	wEncoderID					:WORD := 0; 				(* Encoder ID number *)
	lrTaskCycle					:LREAL := 0.002; 			(* Cycle time of the task which is defined for NC [sec] *)
	bCountDirInv					:BOOL := FALSE;			(* Counting direction inverted if TRUE *)
	udnScalingDenom				:UDINT := 1;	  			(* Denominator for the conversion factor at the conversion of bus data to technical units [INC] *)
	lrScalingNum					:LREAL := 1.0;  			(* Numerator for the conversion factor at the conversion of bus data to technical units [technical units] *)
														(* The technical units dependent on denominator and numerator.*)
	lrModuloFactor 				:LREAL := 360.0; 			(* The "distance" represented by one rotation [technical units] *) 
	dwModuloValue				:DWORD := 0; 			(* Maximum encoder modulo value e.g 1048576 [inc] *)
	etScalingMethod				:ET_ScalingMethod := ET_ScalingMethod_eSMLinear; (* Scaling method: linear or rotary *)
	bSWLimitMaxEn				:BOOL := FALSE;			(* Activation and deactivation of the monitoring of the maximum end position. *)
	lrSWPosLimitMax				:LREAL := 0.0;				(* Location of the maximum end position [technical units] *)
	bSWLimitMinEn 				:BOOL := FALSE;			(* Activation and deactivation of the monitoring of the minimum end position. *)
	lrSWPosLimitMin				:LREAL := 0.0;				(* Location of the minimum end position [technical units] *)

END_STRUCT
END_TYPE

// ---- Data types/Objects/Axis/InternalMC/ST_AXIS_REF_V2.TcDUT
TYPE ST_AXIS_REF_V2 : FB_AXIS_REF_V2;
END_TYPE

// ---- Data types/Objects/EtherCAT Diag/ET_EtherCATDiag.TcDUT
TYPE ET_EtherCATDiag :
(
	ET_EtherCATDiag_eIdle := 0,
	ET_EtherCATDiag_eGetSlaveAdresses,
	ET_EtherCATDiag_eGetSlaveStates,
	ET_EtherCATDiag_eGetTopologyDataLen,
	ET_EtherCATDiag_eGetTopologyData,
	ET_EtherCATDiag_eScanSlaves,
	ET_EtherCATDiag_eGetSlaveIdentity,
	ET_EtherCATDiag_eGetSlaveName,
	ET_EtherCATDiag_eGetScannedSlaveName,
	ET_EtherCATDiag_eDone := 197
);
END_TYPE

// ---- Data types/Objects/EtherCAT Diag/E_EcCommState.TcDUT
TYPE E_EcCommState : (
	eEcState_UNDEFINED 	:= 0,
	eEcState_INIT 		:= 1,
	eEcState_PREOP 		:= 2,
	eEcState_BOOT 		:= 3,
	eEcState_SAFEOP 	:= 4,
	eEcState_OP 		:= 8
);
END_TYPE

// ---- Data types/Objects/EtherCAT Diag/ST_EcMasterDevState.TcDUT
TYPE ST_EcMasterDevState :
STRUCT
	eEcState	 		: E_EcCommState;
	nReserved			: ARRAY [0..2] OF UINT;

	bLinkError			: BOOL;
	bResetRequired		: BOOL;
	bMissFrmRedMode		: BOOL;
	bWatchdogTriggerd	: BOOL;
	bDriverNotFound		: BOOL;
	bResetActive		: BOOL;
	bAtLeastOneNotInOp	: BOOL;
	bDcNotInSync		: BOOL;
END_STRUCT
END_TYPE

// ---- Data types/Objects/EtherCAT Diag/ST_SlaveState.TcDUT
TYPE ST_SlaveState :
STRUCT
	(* slave state *)
	eEcState 		: E_EcCommState;
	nReserved		: UINT;
	bError			: BOOL;
	bInvalidVPRS	: BOOL;
	nReserved2		: UINT;

	(* link state *)
	bNoCommToSlave	: BOOL;
	bLinkError		: BOOL;
	bMissingLink	: BOOL;
	bUnexpectedLink	: BOOL;
	bPortA			: BOOL;
	bPortB			: BOOL;
	bPortC			: BOOL;
	bPortD			: BOOL;
END_STRUCT
END_TYPE

// ---- Data types/Objects/EtherCAT Diag/ST_SlaveStateInfo.TcDUT
TYPE ST_SlaveStateInfo :
STRUCT
	nIndex 			: DINT;
	sName 			: STRING; 		(* name of slave given in System Manager *)
	sType 			: STRING;		(* type of slave, e.g. EK1100*)
	nECAddr 		: UINT;			(* EtherCAT Slave Addr *)
	bDiagData		: BOOL;			(* DiagData in Slave State *)
	stPortCRCErrors	: ST_EcCrcErrorEx;(* Slave CRC-Errors, separate for each Port *)
	nSumCRCErrors	: UDINT;		(* Slave CRC-Errors, sum of all Ports *)
	stState 		: ST_SlaveState;(* EtherCAT State and Link state*)
END_STRUCT
END_TYPE

// ---- Data types/Objects/EtherCAT Diag/ST_SlaveStateInfoScanned.TcDUT
TYPE ST_SlaveStateInfoScanned :
STRUCT
	nIndex 			: DINT;
	sName 			: STRING; 		(* name of slave given in System Manager *)
	sType 			: STRING;		(* type of slave, e.g. EK1100*)
	nECAddr 		: UINT;			(* EtherCAT Slave Addr *)
	bDifferentName	: BOOL;			(* Name of Scanned configuration differs from Configured configuration *)
	bDifferentType	: BOOL;			(* Type Of Scanned configuration differs from Configured configuration *)
	bDifferentAddr	: BOOL;			(* EcAddress of Scanned configuration differs from Configured configuration *)
END_STRUCT
END_TYPE

// ---- Data types/Objects/EtherCAT Diag/ST_TopologyData.TcDUT
TYPE ST_TopologyData :
STRUCT
	iOwnPhysicalAddr 	: UINT;
	iOwnAutoIncAddr		: UINT;
	stPhysicalAddr		: ST_PortAddr;
	stAutoIncAddr		: ST_PortAddr;
	iPortDelay			: ARRAY [0..2] OF UDINT; (* EC_AD, EC_DB, EC_BC *)
	iReserved			: ARRAY [0..7] OF UDINT;
END_STRUCT
END_TYPE

// ---- Data types/Objects/ET_SpindleCtrl/ET_SpindleCtrl.TcDUT
TYPE ET_SpindleCtrl :
(
	ET_SpindleCtrl_eWaitExecute := 0,
	ET_SpindleCtrl_eCtrlEnable := 5,
	ET_SpindleCtrl_eWfCtrlEnabled := 10,
	ET_SpindleCtrl_eSpindleStop := 15,
	ET_SpindleCtrl_eWfSpindleStopped := 20,
	ET_SpindleCtrl_eSpindleRun := 25,
	ET_SpindleCtrl_eWfSpindleRunning := 30,
	ET_SpindleCtrl_eDone := 197,
	ET_SpindleCtrl_eError := 198,
	ET_SpindleCtrl_eNoExecute := 199
);
END_TYPE

// ---- Data types/Objects/FB_Alarm/ET_AlarmType.TcDUT
TYPE ET_AlarmType :
(
	ET_AlarmType_eIdle := 0,
	ET_AlarmType_eFatalError := 1,
	ET_AlarmType_eError := 2,
	ET_AlarmType_eWarning := 3,
	ET_AlarmType_eMessage := 4,
	ET_AlarmType_eHint := 5
);
END_TYPE

// ---- Data types/Objects/FB_Alarm/ST_Alarm.TcDUT
TYPE ST_Alarm :
STRUCT
	bFatalError			:BOOL;				(* Fatal error in group / Fataler Fehler in der Gruppe *)
	bError				:BOOL;				(* Error in group / Fehler in der Gruppe *)
	bWarning			:BOOL;				(* Warning in group / Warnung  in der Gruppe *)
	bMessage			:BOOL;				(* Message in group / Meldung in der Gruppe *)
	bHint				:BOOL;				(* Hint in group / Hint in der Gruppe *)
END_STRUCT
END_TYPE

// ---- Data types/Objects/FB_Alarm/ST_AlarmIn.TcDUT
TYPE ST_AlarmIn :
STRUCT
	arbFatalError			:ARRAY[0..nALARM_MAX_NO] OF ST_AlarmProperties;
	arbError				:ARRAY[0..nALARM_MAX_NO] OF ST_AlarmProperties;
	arbWarning			:ARRAY[0..nALARM_MAX_NO] OF ST_AlarmProperties;
	arbMessage			:ARRAY[0..nALARM_MAX_NO] OF ST_AlarmProperties;
	arbHint				:ARRAY[0..nALARM_MAX_NO] OF ST_AlarmProperties;
END_STRUCT
END_TYPE

// ---- Data types/Objects/FB_Alarm/ST_AlarmOut.TcDUT
TYPE ST_AlarmOut :
STRUCT
	arbFatalError			:ARRAY[0..nALARM_MAX_NO] OF ST_AlarmProperties;
	arbError				:ARRAY[0..nALARM_MAX_NO] OF ST_AlarmProperties;
	arbWarning			:ARRAY[0..nALARM_MAX_NO] OF ST_AlarmProperties;
	arbMessage			:ARRAY[0..nALARM_MAX_NO] OF ST_AlarmProperties;
	arbHint				:ARRAY[0..nALARM_MAX_NO] OF ST_AlarmProperties;
	bFatalError			:BOOL;				(* Fatal error in group / Fataler Fehler in der Gruppe *)
	bError				:BOOL;				(* Error in group / Fehler in der Gruppe *)
	bWarning			:BOOL;				(* Warning in group / Warnung  in der Gruppe *)
	bMessage			:BOOL;				(* Message in group / Meldung in der Gruppe *)
	bHint				:BOOL;				(* Hint in group / Hint in der Gruppe *)
END_STRUCT
END_TYPE

// ---- Data types/Objects/FB_Alarm/ST_AlarmProperties.TcDUT
TYPE ST_AlarmProperties :
STRUCT
	bActive				:BOOL;				(* Alarm on *)
	dtDateTime			:DATE_AND_TIME ;	(* Alarm time stamp *)
	enType				:ET_AlarmType;		(* Alarm type *)
	dnCode				:DINT;				(* Alarm code *)
END_STRUCT
END_TYPE

// ---- Data types/Objects/FB_Alarm/ST_AlarmRef.TcDUT
TYPE ST_AlarmRef :
STRUCT
	stControl					:ST_AlarmOut;
	stManual					:ST_AlarmOut;
	stMaintenance			:ST_AlarmOut;
	stHome					:ST_AlarmOut;
	stAuto					:ST_AlarmOut;
END_STRUCT
END_TYPE

// ---- Data types/Objects/FB_AxisController/ET_AxisGetLimits.TcDUT
TYPE ET_AxisGetLimits :
(
	ET_AxisGetLimits_eWaitExecute := 0,
	ET_AxisGetLimits_eReadVeloMax,
	ET_AxisGetLimits_eWfReadVeloMax,
	ET_AxisGetLimits_eReadAccMax,
	ET_AxisGetLimits_eWfReadAccMax,
	ET_AxisGetLimits_eReadDecMax,
	ET_AxisGetLimits_eWfReadDecMax,
	ET_AxisGetLimits_eReadJerkMax,
	ET_AxisGetLimits_eWfReadJerkMax,
	ET_AxisGetLimits_eReadSoftLimitMax,
	ET_AxisGetLimits_eWfReadSoftLimitMax,
	ET_AxisGetLimits_eReadSoftLimitMin,
	ET_AxisGetLimits_eWfReadSoftLimitMin,
	ET_AxisGetLimits_eDone := 197,
	ET_AxisGetLimits_eError := 198,
	ET_AxisGetLimits_eNoExecute := 199
);
END_TYPE

// ---- Data types/Objects/FB_AxisController/ET_AxisSetLimits.TcDUT
TYPE ET_AxisSetLimits :
(
	ET_AxisSetLimits_eWaitExecute := 0,
	ET_AxisSetLimits_eSetReferenceSystem,
	ET_AxisSetLimits_eWfSetReferenceSystem,
	ET_AxisSetLimits_eSetPositionBias,
	ET_AxisSetLimits_eWfSetPositionBias,
	ET_AxisSetLimits_eSetLimitPos,
	ET_AxisSetLimits_eWfSetLimitPos,
	ET_AxisSetLimits_eSetLimitNeg,
	ET_AxisSetLimits_eWfSetLimitNeg,
	ET_AxisSetLimits_eEnableLimitPos,
	ET_AxisSetLimits_eWfEnableLimitPos,
	ET_AxisSetLimits_eEnableLimitNeg,
	ET_AxisSetLimits_eWfEnableLimitNeg,
	ET_AxisSetLimits_eEnablePosLagMonitoring,
	ET_AxisSetLimits_eWfEnablePosLagMonitoring,
	ET_AxisSetLimits_eDone := 197,
	ET_AxisSetLimits_eError := 198,
	ET_AxisSetLimits_eNoExecute := 199
);
END_TYPE

// ---- Data types/Objects/FB_AxisController/ET_STOEBER_AxisGetLimitsTc2.TcDUT
TYPE ET_STOEBER_AxisGetLimitsTc2 :
(
	ET_STOEBER_AxisGetLimits_eWaitExecute := 0,
	ET_STOEBER_AxisGetLimits_eDecimalDigits,
	ET_STOEBER_AxisGetLimits_eScalingDenom,
	ET_STOEBER_AxisGetLimits_eScalingNum,
	ET_STOEBER_AxisGetLimits_eDone := 197,
	ET_STOEBER_AxisGetLimits_eError := 198,
	ET_STOEBER_AxisGetLimits_eNoExecute := 199
);
END_TYPE

// ---- Data types/Objects/FB_AxisController/ET_STOEBER_AxisSetLimitsTc2.TcDUT
TYPE ET_STOEBER_AxisSetLimitsTc2 :
(
	ET_STOEBER_AxisSetLimits_eWaitExecute := 0,
	ET_STOEBER_AxisSetLimits_eSetLimitPos,
	ET_STOEBER_AxisSetLimits_eSetLimitNeg,
	ET_STOEBER_AxisSetLimits_eSetJogVelo,
	ET_STOEBER_AxisSetLimits_eSetJogAcc,
	ET_STOEBER_AxisSetLimits_eSetJogDec,
	ET_STOEBER_AxisSetLimits_eSetJogJerk,
	ET_STOEBER_AxisSetLimits_eDone := 197,
	ET_STOEBER_AxisSetLimits_eError := 198,
	ET_STOEBER_AxisSetLimits_eNoExecute := 199
);
END_TYPE

// ---- Data types/Objects/FB_AxisMoveManual/ET_AxisMoveManualSetLimits.TcDUT
TYPE ET_AxisMoveManualSetLimits :
(
	ET_AxisMoveManualSetLimits_eWaitExecute := 0,
	ET_AxisMoveManualSetLimits_eSetVelo := 5,
	ET_AxisMoveManualSetLimits_eWfSetVelo := 10,
	ET_AxisMoveManualSetLimits_eDone := 197,
	ET_AxisMoveManualSetLimits_eError := 198,
	ET_AxisMoveManualSetLimits_eNoExecute := 199
);
END_TYPE

// ---- Data types/Objects/FB_Blinker/ST_Blinker.TcDUT
TYPE ST_Blinker :
STRUCT	
	Q0					:BOOL; 						(* Divider output / 2 *)
	Q1					:BOOL; 						(* Divider output / 4 *)
	Q2					:BOOL; 						(* Divider output / 8 *)
	Q3					:BOOL; 						(* Divider output / 16 *)
	Q4					:BOOL; 						(* Divider output / 32 *)
	Q5					:BOOL; 						(* Divider output / 64 *)
	Q6					:BOOL; 						(* Divider output / 128 *)
	Q7					:BOOL; 						(* Divider output / 256 *)
END_STRUCT
END_TYPE

// ---- Data types/Objects/FB_CalcContour/ET_ContourType.TcDUT
TYPE ET_ContourType :
(
	ET_ContourType_eNone := 0,
	ET_ContourType_eCircle := 1,
	ET_ContourType_eEllipse := 2,
	ET_ContourType_eSquare := 3
);
END_TYPE

// ---- Data types/Objects/FB_CfgAxisInExt3DGroup/ET_CfgAxisInExt3DGroup.TcDUT
TYPE ET_CfgAxisInExt3DGroup :
(
	ET_CfgAxisInExt3DGrp_eWaitExecute := 0,
	ET_CfgAxisInExt3DGrp_eReadExt3DAxisIds := 5,
	ET_CfgAxisInExt3DGrp_eDone := 197,
	ET_CfgAxisInExt3DGrp_eError := 198,
	ET_CfgAxisInExt3DGrp_eNoExecute := 199
);
END_TYPE

// ---- Data types/Objects/FB_DistanceCounter/ST_DistanceCounter.TcDUT
TYPE ST_DistanceCounter :
STRUCT
	lrAllOverDistance					:LREAL; 							(* All over counter distance *)
	lrAfterResetDistance				:LREAL; 							(* Counter distance since last reset *)
END_STRUCT
END_TYPE

// ---- Data types/Objects/FB_EL3312/ET_EL3312ThermocoupleTyp.TcDUT
TYPE ET_EL3312ThermocoupleTyp :
(
	ET_EL3312ThermocoupleTyp_eK := 0,				(* Typ: K -200°C bis 1370°C *)
	ET_EL3312ThermocoupleTyp_eJ := 1,				(* Typ: J -100°C bis 1200°C *)
	ET_EL3312ThermocoupleTyp_eL := 2,				(* Typ: L 0°C bis 900°C *)
	ET_EL3312ThermocoupleTyp_eE := 3,				(* Typ: E -100°C bis 1000°C *)
	ET_EL3312ThermocoupleTyp_eT := 4,				(* Typ: T -200°C bis 400°C *)
	ET_EL3312ThermocoupleTyp_eN := 5,				(* Typ: N -100°C bis 1300°C *)
	ET_EL3312ThermocoupleTyp_eU := 6,				(* Typ: U 0°C bis 600°C *)
	ET_EL3312ThermocoupleTyp_eB := 7,				(* Typ: B 600°C bis 1800°C *)
	ET_EL3312ThermocoupleTyp_eR := 8,				(* Typ: R 0°C bis 1767°C *)
	ET_EL3312ThermocoupleTyp_eS := 9,				(* Typ: S 0°C bis 1760°C *)
	ET_EL3312ThermocoupleTyp_eC := 10,				(* Typ: C 0°C bis 2320°C *)
	ET_EL3312ThermocoupleTyp_e30mV := 100,			(* +/-30 mV (1uV resolution) *)
	ET_EL3312ThermocoupleTyp_e60mV := 101,			(* +/-60 mV (2uV resolution) *)
	ET_EL3312ThermocoupleTyp_e75mV := 102,			(* +/-75 mV (4uV resolution) *)
	ET_EL3312ThermocoupleTyp_eNoConn := 999		(* No connected *)
);
END_TYPE

// ---- Data types/Objects/FB_EL3312/ST_EL3312ChannelState.TcDUT
TYPE ST_EL3312ChannelState :
STRUCT
	bUnderrange				:BOOL;			(* State underrange *)
	bOverrange				:BOOL;			(* State overrange *)
	byLimit1					:BYTE;			(* State limit 1 *)
	byLimit2 					:BYTE;			(* State limit 2 *)
	bError 					:BOOL;			(* State error *)
	bState 					:BOOL;			(* State *)
	bToggle					:BOOL;			(* TxPDO Toggle *)
END_STRUCT
END_TYPE

// ---- Data types/Objects/FB_EL3312/ST_EL3312CoeInfo.TcDUT
TYPE ST_EL3312CoeInfo :
STRUCT
	bEnableUserScale 			:BOOL := FALSE;
	bEnableFilter 					:BOOL := FALSE;
	bEnableLimit1 				:BOOL := FALSE;
	bEnableLimit2 				:BOOL := FALSE;
	bEnableUserCalibration 		:BOOL := FALSE;
	bEnableVendorCalibration 		:BOOL := TRUE;
	dwColdjunctionCompensation 	:DWORD := 0;
	nUserScaleOffset 				:INT := 0;
	dnUserScaleGain 				:DINT := 65536;
	nLimit1 						:INT := 0;
	nLimit2 						:INT := 0;
	dwFilterSettings 				:DWORD := 0;
	nUserCalibrationOffset 			:INT := 0;
	unUserCalibrationGain 			:UINT := 65535;
	dwTCElement 				:DWORD := 0;
END_STRUCT
END_TYPE

// ---- Data types/Objects/FB_EL3312/ST_EL3312CoeReadData.TcDUT
TYPE ST_EL3312CoeReadData :
STRUCT
	wIdx: WORD;
	bySubIdx: BYTE;
	bReadOK: BOOL;
	dwData: DWORD;
	nSize: UDINT;
END_STRUCT
END_TYPE

// ---- Data types/Objects/FB_EL3312/ST_EL3312CoeWriteData.TcDUT
TYPE ST_EL3312CoeWriteData :
STRUCT
	wIdx: WORD;
	bySubIdx: BYTE;
	bWriteOK: BOOL;
	dwData: DWORD;
	nSize: UDINT;
END_STRUCT
END_TYPE

// ---- Data types/Objects/FB_EL3351/ST_EL3351ChannelState.TcDUT
TYPE ST_EL3351ChannelState :
STRUCT
	bUnderrange				:BOOL;			(* State underrange *)
	bOverrangerange			:BOOL;			(* State overrangerange *)
	bError 					:BOOL;			(* State error *)
	bState 					:BOOL;			(* State *)
	bToggle					:BOOL;			(* TxPDO Toggle *)
END_STRUCT
END_TYPE

// ---- Data types/Objects/FB_EL3351/ST_EL3351CoeInfo.TcDUT
TYPE ST_EL3351CoeInfo :
STRUCT
	bEnableUserScale: BOOL:= 0;
	diUserScaleOffset: DINT:= 0;
	diUserScaleGain: DINT:= 65536;
	dwFilterSettings: DWORD:= 2;

	bEnableUserScaleIndex8010: BOOL:= 0;
	dnUserScaleOffsetIndex8010: DINT:= 0;
	dnUserScaleGainIndex8010: DINT:= 65536;
END_STRUCT
END_TYPE

// ---- Data types/Objects/FB_EL3351/ST_EL3351CoeReadData.TcDUT
TYPE ST_EL3351CoeReadData :
STRUCT
	wIdx: WORD;
	bySubIdx: BYTE;
	bReadOK: BOOL;
	nData: UDINT;
	nSize: UDINT;
END_STRUCT
END_TYPE

// ---- Data types/Objects/FB_EL3351/ST_EL3351CoeWriteData.TcDUT
TYPE ST_EL3351CoeWriteData :
STRUCT
	wIdx: WORD;
	bySubIdx: BYTE;
	bWriteOK: BOOL;
	nData: DWORD;
	nSize: UDINT;
END_STRUCT
END_TYPE

// ---- Data types/Objects/FB_EL3356/ST_EL3356ChannelCtrl.TcDUT
TYPE ST_EL3356ChannelCtrl :
STRUCT
	bStartCalibration			:BOOL;			(* Ctrl start calibration *)
	bDisableCalibration		:BOOL;			(* Ctrl disable calibration *)
	bInputFreeze				:BOOL;			(* Ctrl input freeze *)
	bTare					:BOOL;			(* Ctrl tare *)
END_STRUCT
END_TYPE

// ---- Data types/Objects/FB_EL3356/ST_EL3356ChannelState.TcDUT
TYPE ST_EL3356ChannelState :
STRUCT
	bOverrange				:BOOL;			(* State Overrange *)
	bDataInvalid				:BOOL;			(* State Data invalid *)
	bError 					:BOOL;			(* State error *)
	bCalibrationInProgress 	:BOOL;			(* State calibration in progress *)
	bSteadyState 			:BOOL;			(* Stady state *)
	bSyncError				:BOOL;			(* Sync error *)
	bToggle					:BOOL;			(* TxPDO Toggle *)
END_STRUCT
END_TYPE

// ---- Data types/Objects/FB_EL3356/ST_EL3356CoeInfo.TcDUT
TYPE ST_EL3356CoeInfo :
STRUCT
	bEnableFilter							:BOOL:= TRUE;
	bEnableUserScale					:BOOL:= TRUE;
	dwFilterSettings						:DWORD:= 0;
	rGain								:REAL:= 1.0;
	rTara								:REAL:= 0.0;
	rRatedOutput							:REAL:= 2.0;
	rNominalLoad						:REAL:= 5.0;
	rZeroBalance							:REAL:= 0.0;
	rGravityOfEarth						:REAL:= 9.806650;
	rScaleFactor							:REAL:= 1000.0;
	rReferenceLoad						:REAL:= 5.0;
	bEnableUserScaleIndex8010			:BOOL:= FALSE;
	dnUserScaleOffsetIndex8010			:DINT:= 0;
	dnUserScaleGainIndex8010				:DINT:= 65536;
	dwFilterSettingsIndex8010				:DWORD:= 0;
END_STRUCT
END_TYPE

// ---- Data types/Objects/FB_EL3356/ST_EL3356CoeReadData.TcDUT
TYPE ST_EL3356CoeReadData :
STRUCT
	wIdx: WORD;
	bySubIdx: BYTE;
	bReadOK: BOOL;
	dwData: DWORD;
	nSize: UDINT;
END_STRUCT
END_TYPE

// ---- Data types/Objects/FB_EL3356/ST_EL3356CoeWriteData.TcDUT
TYPE ST_EL3356CoeWriteData :
STRUCT
	wIdx: WORD;
	bySubIdx: BYTE;
	bWriteOK: BOOL;
	dwData: DWORD;
	nSize: UDINT;
END_STRUCT
END_TYPE

// ---- Data types/Objects/FB_ExtSetPoint/ET_MoveExtState.TcDUT
TYPE ET_MoveExtState :
(
	ET_MoveExtState_eWaitExecute := 0,
	ET_MoveExtState_eEnableExtSetPointGenerator := 5,
	ET_MoveExtState_eDisableExtSetPointGenerator := 10,
	ET_MoveExtState_eDone := 197,
	ET_MoveExtState_eError := 198,
	ET_MoveExtState_eNoExecute := 199
);
END_TYPE

// ---- Data types/Objects/FB_ExtTrajPos/ET_CalcExtTrajState.TcDUT
TYPE ET_CalcExtTrajState :
(
	ET_CalcExtTrajState_eWaitExecute := 0,
	ET_CalcExtTrajState_eCalcTrajPos := 5,
	ET_CalcExtTrajState_eDone := 197,
	ET_CalcExtTrajState_eError := 198,
	ET_CalcExtTrajState_eNoExecute := 199
);
END_TYPE

// ---- Data types/Objects/FB_ItpReadRParams/ET_ItpReadRParams.TcDUT
TYPE ET_ItpReadRParams :
(
	ET_ItpReadRParams_eWaitExecute := 0,
	ET_ItpReadRParams_eReadRParams := 5,
	ET_ItpReadRParams_eDone := 197,
	ET_ItpReadRParams_eError := 198,
	ET_ItpReadRParams_eNoExecute := 199
);
END_TYPE

// ---- Data types/Objects/FB_ItpWriteRParams/ET_ItpWriteRParams.TcDUT
TYPE ET_ItpWriteRParams :
(
	ET_ItpWriteRParams_eWaitExecute := 0,
	ET_ItpWriteRParams_eWriteRParams := 5,
	ET_ItpWriteRParams_eDone := 197,
	ET_ItpWriteRParams_eError := 198,
	ET_ItpWriteRParams_eNoExecute := 199
);
END_TYPE

// ---- Data types/Objects/FB_KL600x/ET_KL600xInit.TcDUT
TYPE ET_KL600xInit :
(
	ET_KL600xInit_eInit := 0,
	ET_KL600xInit_eChkSettings,
	ET_KL600xInit_eWriteEnableRTSCTS,
	ET_KL600xInit_eWriteBaudRate,
	ET_KL600xInit_eWriteDataFrame,
	ET_KL600xInit_eDone := 197,
	ET_KL600xInit_eError := 198,
	ET_KL600xInit_eNoExecute := 199
);
END_TYPE

// ---- Data types/Objects/FB_KL600x/ET_KL600xSend.TcDUT
TYPE ET_KL600xSend :
(
	ET_KL600xSend_eInit := 0,
	ET_KL600xSend_eSend,
	ET_KL600xSend_eDone := 197,
	ET_KL600xSend_eError := 198,
	ET_KL600xSend_eNoExecute := 199
);
END_TYPE

// ---- Data types/Objects/FB_KL600x/ST_KL600xData.TcDUT
TYPE ST_KL600xData :
STRUCT
	sDateTime			:STRING;
	sData				:STRING;
END_STRUCT
END_TYPE

// ---- Data types/Objects/FB_LoadFromFile/ET_LoadFromFile.TcDUT

TYPE ET_LoadFromFile :
(
	ET_LoadFromFile_eWaitExecute := 0,
	ET_LoadFromFile_eFileName,
	ET_LoadFromFile_eChkFileExist,
	ET_LoadFromFile_eFileOpen,
	ET_LoadFromFile_eChkFileOpen,
	ET_LoadFromFile_eReadData,
	ET_LoadFromFile_eChkReadData,
	ET_LoadFromFile_eFileClose,
	ET_LoadFromFile_eChkFileClose,
	ET_LoadFromFile_eDone := 197,
	ET_LoadFromFile_eError := 198,
	ET_LoadFromFile_eNoExecute := 199
);
END_TYPE

// ---- Data types/Objects/FB_Logger/ST_Logger.TcDUT
TYPE ST_Logger :
STRUCT
	arstLoggerWaitInterrupt					:ARRAY[1..unLOG_BEFOR_MAX_NO] OF ST_LoggerVar;
	arstLoggerDuringInterrupt				:ARRAY[1..unLOG_DURING_MAX_NO] OF ST_LoggerVar;
	arstLoggerAfterInterrupt					:ARRAY[1..unLOG_AFTER_MAX_NO] OF ST_LoggerVar;
END_STRUCT
END_TYPE

// ---- Data types/Objects/FB_Logger/ST_LoggerVar.TcDUT
TYPE ST_LoggerVar :
STRUCT
	udnCycleNo		:UDINT;
	sTimeStamp		:STRING(15);			(* Alarm time stamp *)
	arsLogVars		:ARRAY[1..unNUM_OF_LOG_VAR] OF STRING(10);
END_STRUCT
END_TYPE

// ---- Data types/Objects/FB_ModeSelector/ET_MachineMode.TcDUT
(* Machine operating mode *)
TYPE ET_MachineMode :
(
	ET_MachineMode_eUndefined := 0,
	ET_MachineMode_eAutomatic := 1,
	ET_MachineMode_eCycle := 2,
	ET_MachineMode_eStepping := 3,
	ET_MachineMode_eHome := 4,
	ET_MachineMode_eManual := 5,
	ET_MachineMode_eMaintenance := 6,
	ET_MachineMode_eDryRun := 7,
	ET_MachineMode_eMDI := 8,
	ET_MachineMode_eIdle := 10
);
END_TYPE

// ---- Data types/Objects/FB_ModeSelector/ET_MachineState.TcDUT
(* Machine state *)
TYPE ET_MachineState :
(
	ET_MachineState_eUndefined := 0,
	ET_MachineState_eAutoExe := 1,
	ET_MachineState_eAutoSteppingExe := 2,
	ET_MachineState_eAutoSteppingNoExe := 3,
	ET_MachineState_eHomeExe := 4,
	ET_MachineState_eHomeRefExe := 5,
	ET_MachineState_eMaintenanceExe := 6,
	ET_MachineState_eIdle := 10
) ;
END_TYPE

// ---- Data types/Objects/FB_RampDirector/ET_RampGenerator.TcDUT
TYPE ET_RampGenerator :
(
	ET_RampGenerator_eWaitExecute := 0,
	ET_RampGenerator_eRunning := 5,
	ET_RampGenerator_eWaiting := 10,
	ET_RampGenerator_eDone := 197,
	ET_RampGenerator_eError := 198,
	ET_RampGenerator_eNotExecute := 199
);
END_TYPE

// ---- Data types/Objects/FB_SpindlePreheat/ET_SpindlePreheat.TcDUT
TYPE ET_SpindlePreheat :
(
	ET_SpindlePreheat_eWaitExecute := 0,
	ET_SpindlePreheat_eStartNewSpindle := 5,
	ET_SpindlePreheat_eStartDailyPreheat := 10,
	ET_SpindlePreheat_eStartSpindle := 15,
	ET_SpindlePreheat_eWfStartSpindle := 20,
	ET_SpindlePreheat_eWfStartSpindleProc := 25,
	ET_SpindlePreheat_eSpindleStop := 30,
	ET_SpindlePreheat_eWfSpindleStopped := 35,
	ET_SpindlePreheat_eDone := 197,
	ET_SpindlePreheat_eError := 198,
	ET_SpindlePreheat_eNoExecute := 199
);
END_TYPE

// ---- Data types/Objects/FB_SpindlePreheat/ST_SpindlePreheat.TcDUT
TYPE ST_SpindlePreheat :
STRUCT
	dwOverride				:DWORD;			(* Override is percent of total speed of spindle. The range of override is from 0%  to 100 %  of rated speed.*)
	tDuration					:TIME;				(* Duration time for current phase *)
	dwSpeedRpm			:DWORD;			(* Current speed RPM - Read Only *)
	otstDuration				:OTSTRUCT;			(* Duration time in OTSTRUCT - Read Only*)
END_STRUCT
END_TYPE

// ---- Data types/Objects/FB_TimeHoursCounter/ST_TimeHoursCounter.TcDUT
TYPE ST_TimeHoursCounter :
STRUCT
	lrAllOverHours					:LREAL; 							(* All over counter hours *)
	lrAfterResetHours					:LREAL; 							(* Counter hours since last reset *)
END_STRUCT
END_TYPE

// ---- Data types/Objects/FB_Timer/ST_DateTime.TcDUT
TYPE ST_DateTime :
STRUCT
	sDate						:STRING;					(* Current data *)
	sTime						:STRING;					(* Current time *)
	sTimeEx						:STRING;					(* Current time extend *)
	sDateTime					:STRING;					(* Current data and time *)
	dtDateTime					:DATE_AND_TIME;				(* Current data and time *)
	sDateTimeEx					:STRING;					(* Current data and time extend *)
	dtDateTimeEx				:DATE_AND_TIME;				(* Current data and time extend *)
END_STRUCT
END_TYPE

// ---- Data types/Objects/FB_Timer/ST_Time.TcDUT
TYPE ST_Time :
STRUCT
	dwSec				:DWORD; 						(* Time in 1 [s] *)
	dwDeciSec			:DWORD; 						(* Time in deci 0.1 [s] *)
	dwCentiSec			:DWORD; 						(* Time in centi 0.01 [s] *)
	dwMiliSec			:DWORD; 						(* Time in mili 0.001 [s] *)
END_STRUCT
END_TYPE

// ---- Data types/Objects/FB_ToolStorage/ET_ToolStatus.TcDUT
TYPE ET_ToolStatus :
(
	ET_ToolStatus_eOk,
	ET_ToolStatus_eNOk,
	ET_ToolStatus_eLifettimeExceeded
);
END_TYPE

// ---- Data types/Objects/FB_ToolStorage/ET_ToolStorage.TcDUT
TYPE ET_ToolStorage :
(
	ET_ToolStorage_eWaitExecute := 0,
	ET_ToolStorage_eGetNewToolNest,
	ET_ToolStorage_eGetOldToolNest,
	ET_ToolStorage_eChkToolPlace,
	ET_ToolStorage_eChkToolPickUp,
	ET_ToolStorage_eDone := 197,
	ET_ToolStorage_eError := 198,
	ET_ToolStorage_eNoExecute := 199
);
END_TYPE

// ---- Data types/Objects/FB_Traceability/ST_Traceability.TcDUT
TYPE ST_Traceability :
STRUCT
	sDateTime				:STRING(15);
	stSettings				:ST_TraceabilitySettings;
	arstData					:ARRAY[1..udnTraceSampleMax,1..udnTraceDataMax] OF ST_TraceabilityData;
END_STRUCT
END_TYPE

// ---- Data types/Objects/FB_Traceability/ST_TraceabilityData.TcDUT
TYPE ST_TraceabilityData :
STRUCT
	sName					:STRING(15);
	sValue					:STRING(15);
	sUnit					:STRING(5);
END_STRUCT
END_TYPE

// ---- Data types/Objects/FB_Traceability/ST_TraceabilitySettings.TcDUT
TYPE ST_TraceabilitySettings :
STRUCT
	sPath								:STRING;						(* Path to file e.g. 'c:\', Hard Disk\ *)
	sFileName							:STRING(20);						(* Name of file *)
	sFileExtension						:STRING(5);						(* File extension  *)
END_STRUCT
END_TYPE

// ---- Data types/Objects/Fieldbus/ST_FieldbusStatus.TcDUT
TYPE ST_FieldbusStatus :
STRUCT
	wFrmXWcState				:WORD; (* link to task related ethercat frame state FrmXWcState *)
	nMasterDeviceId				:UINT;
	nMasterSlaveCount			:UINT;
	nMasterDevState				:UINT;
	arrMasterNetId				:T_AmsNetIdArr;
	nMasterSlaveCountCfg			:UINT;
END_STRUCT
END_TYPE

// ---- Data types/Objects/Gefran/ET_GFX4IR.TcDUT
TYPE ET_GFX4IR :
(
	ET_GFX4IRState_eWaitExecute := 0,
	ET_GFX4IRState_eCtrlOn,
	ET_GFX4IRState_eCtrlOff,
	ET_GFX4IRState_eDone := 197,
	ET_GFX4IRState_eError := 198,
	ET_GFX4IRState_eNoExecute := 199
);
END_TYPE

// ---- Data types/Objects/Gefran/ST_GFX4IRTOPLC.TcDUT
TYPE ST_GFX4IRTOPLC:
STRUCT
	nProcessVariable			:INT;
	wControllerStatus			:WORD;
	nOutputPower				:INT;
	wAmmeterInputOn			:WORD;
END_STRUCT
END_TYPE

// ---- Data types/Objects/Gefran/ST_GFX4IR_REF.TcDUT
TYPE ST_GFX4IR_REF : FB_GFX4IR_REF;
END_TYPE

// ---- Data types/Objects/Gefran/ST_PLCTOGFX4IR.TcDUT
TYPE ST_PLCTOGFX4IR :
STRUCT
	nLocalSetPoint			:INT;
	nManualOutput			:WORD;
	wControllerStatus			:WORD;
END_STRUCT
END_TYPE

// ---- Data types/Objects/Leister/ET_LeisterExtruder.TcDUT
TYPE ET_LeisterExtruder :
(
	ET_LeisterExtruder_eWaitExecute := 0,
	ET_LeisterExtruder_eStartExtruder,
	ET_LeisterExtruder_eStopExtruder,
	ET_LeisterExtruder_eWfHeaterReady,
	ET_LeisterExtruder_eDone := 197,
	ET_LeisterExtruder_eError := 198,
	ET_LeisterExtruder_eNoExecute := 199
);
END_TYPE

// ---- Data types/Objects/Leister/ET_LeisterHeater.TcDUT
TYPE ET_LeisterHeater :
(
	ET_LeisterHeater_eWaitExecute := 0,
	ET_LeisterHeater_eStartHeater,
	ET_LeisterHeater_eStopHeater,
	ET_LeisterHeater_eDone := 197,
	ET_LeisterHeater_eError := 198,
	ET_LeisterHeater_eNoExecute := 199
);
END_TYPE

// ---- Data types/Objects/Leister/ST_LEISTERTOPLC.TcDUT
TYPE ST_LEISTERTOPLC :
STRUCT
	arbyInput				:ARRAY[0..63] OF BYTE;
END_STRUCT
END_TYPE

// ---- Data types/Objects/Leister/ST_LEISTER_REF.TcDUT
TYPE ST_LEISTER_REF : FB_LEISTER_EXTRUDER_REF;
END_TYPE

// ---- Data types/Objects/Leister/ST_PLCTOLEISTER.TcDUT
TYPE ST_PLCTOLEISTER :
STRUCT
	arbyOutput				:ARRAY[0..63] OF BYTE;
END_STRUCT
END_TYPE

// ---- Data types/Objects/Munsch/ET_MunschExtruder.TcDUT
TYPE ET_MunschExtruder :
(
	ET_MunschExtruder_eWaitExecute := 0,
	ET_MunschExtruder_eChkInterface,
	ET_MunschExtruder_eSetCMD,
	ET_MunschExtruder_eSetMaterialTemp,
	ET_MunschExtruder_eSetAirTemp,
	ET_MunschExtruder_eExecuteCMD,
	ET_MunschExtruder_eSetREQ,
	ET_MunschExtruder_eExecuteREQ,
	ET_MunschExtruder_eDone := 197,
	ET_MunschExtruder_eError := 198,
	ET_MunschExtruder_eNoExecute := 199
);
END_TYPE

// ---- Data types/Objects/Munsch/ET_MUNSCH_CMD.TcDUT
(* Munsch command *)
TYPE ET_MUNSCH_CMD :
(
	ET_MUNSCH_CMD_NOCMD := 0,
	ET_MUNSCH_CMD_STARTHEAT := 1,
	ET_MUNSCH_CMD_STOPHEAT := 2,
	ET_MUNSCH_CMD_REQHEATSTATUS := 3,
	ET_MUNSCH_CMD_STARTEXTRUDER := 5,
	ET_MUNSCH_CMD_STOPEXTRUDER := 6,
	ET_MUNSCH_CMD_REQEXTRUDERSTATUS := 7,
	ET_MUNSCH_CMD_SETMATERIALTEMP := 9,
	ET_MUNSCH_CMD_REQMATERIALREFTEMP := 10,
	ET_MUNSCH_CMD_REQMATERIALACTTEMP := 11,
	ET_MUNSCH_CMD_SETAIRTEMP := 13,
	ET_MUNSCH_CMD_REQAIRREFTEMP := 14,
	ET_MUNSCH_CMD_REQAIRACTTEMP := 15,
	ET_MUNSCH_CMD_REQSTATUS := 20

);
END_TYPE

// ---- Data types/Objects/Munsch/ET_MUNSCH_RES.TcDUT
(* Munsch response *)
TYPE ET_MUNSCH_RES :
(
	ET_MUNSCH_RES_NOCMD := 0,
	ET_MUNSCH_RES_STARTHEAT := 1,
	ET_MUNSCH_RES_STOPHEAT := 2,
	ET_MUNSCH_RES_ACKHEATSTATUSON := 3,
	ET_MUNSCH_RES_ACKHEATSTATUSOFF := 4,
	ET_MUNSCH_RES_STARTEXTRUDER := 5,
	ET_MUNSCH_RES_STOPEXTRUDER := 6,
	ET_MUNSCH_RES_ACKEXTRUDERSTATUSON := 7,
	ET_MUNSCH_RES_ACKEXTRUDERSTATUSOFF := 8,
	ET_MUNSCH_RES_SETMATERIALTEMP := 9,
	ET_MUNSCH_RES_REQMATERIALREFTEMP := 10,
	ET_MUNSCH_RES_REQMATERIALACTTEMP := 11,
	ET_MUNSCH_RES_SETAIRTEMP := 13,
	ET_MUNSCH_RES_REQAIRREFTEMP := 14,
	ET_MUNSCH_RES_REQAIRACTTEMP := 15,
	ET_MUNSCH_RES_REQSTATUSHEATING := 17,
	ET_MUNSCH_RES_REQSTATUSHEATED := 18,
	ET_MUNSCH_RES_REQSTATUSERROR := 19,
	ET_MUNSCH_RES_CMDERROR := 21

);
END_TYPE

// ---- Data types/Objects/Munsch/ST_MUNSCH_CMD_Data.TcDUT
TYPE ST_MUNSCH_CMD_Data :
STRUCT
	nMaterialTemp				:INT := 0;				(* Material temperatur. unsMaterialTemp is the temperature in °C added to 160 °C. The range is 0 (160 °C) to 240 (400 °C) *)
	nAirTemp					:INT := 0;				(* Air temperatur. unsAirTemp is the temperature in °C added to 160 °C. The range is 0 (160 °C) to 240 (400 °C) *)
	etCommand					:ET_MUNSCH_CMD;
END_STRUCT
END_TYPE

// ---- Data types/Objects/Munsch/ST_MUNSCH_REF.TcDUT
TYPE ST_MUNSCH_REF : FB_MUNSCH_EXTRUDER_REF;
END_TYPE

// ---- Data types/Objects/Munsch/ST_MUNSCH_RES_Data.TcDUT
TYPE ST_MUNSCH_RES_Data :
STRUCT
	nMaterialRefTemp			:INT := 0;				(* Material referenc temperatur. unsMaterialTemp is the temperature in °C added to 160 °C. The range is 0 (160 °C) to 240 (400 °C) *)
	nMaterialActTemp				:INT := 0;				(* Material referenc temperatur. unsMaterialTemp is the temperature in °C added to 160 °C. The range is 0 (160 °C) to 240 (400 °C) *)
	nAirRefTemp					:INT := 0;				(* Air current temperatur. unsAirTemp is the temperature in °C added to 160 °C. The range is 0 (160 °C) to 240 (400 °C) *)
	nAirActTemp					:INT := 0;				(* Air current temperatur. unsAirTemp is the temperature in °C added to 160 °C. The range is 0 (160 °C) to 240 (400 °C) *)
	etResponse					:ET_MUNSCH_RES;
END_STRUCT
END_TYPE

// ---- Data types/Objects/Periphery/ST_PERIPHERYTOPLC.TcDUT
TYPE ST_PERIPHERYTOPLC :
STRUCT

END_STRUCT
END_TYPE

// ---- Data types/Objects/Periphery/ST_PERIPHERY_REF.TcDUT
TYPE ST_PERIPHERY_REF : FB_PERIPHERY_REF;
END_TYPE

// ---- Data types/Objects/Periphery/ST_PLCTOPERIPHERY.TcDUT
TYPE ST_PLCTOPERIPHERY :
STRUCT

	bAllDoorsLocked						:BOOL;						(* IN - All Doors Locked / Alle Türen geschlossen  *)
	bExtStart								:BOOL;						(* IN - External start  *)

	bMachineError						:BOOL;						(* IN - Machine has fault. *)
	bMachineStandstill					:BOOL;						(* IN - Machine standstill. *)
	bMachineReady						:BOOL;						(* IN - Machine ready. *)

	nPrgNoSideA							:INT;						(* IN - Program on side A *)
	nPrgNoSideB							:INT;						(* IN - Program on side B *)
END_STRUCT
END_TYPE

// ---- Data types/Objects/Robot/KUKA/ET_KukaStart.TcDUT
TYPE ET_KukaStart :
(
	ET_KukaStart_eWaitExecute := 0,
	ET_KukaStart_eExtStart,
	ET_KukaStart_eWfInHome,
	ET_KukaStart_eWfPgNoReq,
	ET_KukaStart_ePgNoParity,
	ET_KukaStart_ePgNoValid,
	ET_KukaStart_eWfProgFinish,
	ET_KukaStart_eDone := 197,
	ET_KukaStart_eError := 198,
	ET_KukaStart_eNoExecute := 199
);
END_TYPE

// ---- Data types/Objects/Robot/KUKA/ST_KUKATOPLC.TcDUT
TYPE ST_KUKATOPLC :
STRUCT
	bStopMess						:BOOL;						(* $OUT[1010] - Any message occurring which requires the robot to be stopped / Störung Roboter *)
	bPgNoReq						:BOOL;						(* $OUT[33] - A change of signal requests the higher-level controller to send a program number / PGNO Req-Signalwechsel fordert Leitrechner Programmnr. zu senden *)
	bApplRun						:BOOL;						(* $OUT[34] - Program is currently being executed / TRUE wenn Programm abgearbeitet wird *)
	bPeriRdy						:BOOL;						(* $OUT[1012] - Robot drives are switched on / TRUE wenn Roboterantriebe eingeschaltet *)
	bAlarmStop						:BOOL;						(* $OUT[1013] - Emergency stop / Not Aus *)
	bUserSafe						:BOOL;						(* $OUT[1011] - If the safety fence monitoring switch is opened (AUT mode) or an enabling switch is released (T1 or T2 mode). / Abfrage Schutzgitter(Auto)/Zustimmungsschalter(Test) *)
	bT1								:BOOL;						(* $OUT[993] - Operating mode T1 / Betriebsart T1 *)
	bT2								:BOOL;						(* $OUT[994] - Operating mode T2/ Betriebsart T2 *)
	bAut								:BOOL;						(* $OUT[995] - Operating mode Aut / Betriebsart Aut *)
	bExt								:BOOL;						(* $OUT[996] - Operating mode Ext / Betriebsart Ext *)
	bOnPath							:BOOL;						(* $OUT[997] - Set as long as the robot stays on its programmed path / TRUE solange sich Rob. auf programmierten Bahn befindet *)
	bProAct							:BOOL;						(* $OUT[1021] - Whenever a process is active / Programmbearbeitung aktiv *)
	bInHome							:BOOL;						(* $OUT[1000] - Whether or not the robot is in its HOME position  / In Home Position *)
	arbInHome						:ARRAY[1..5] OF BOOL;		(* $OUT[1003..1007] - Whether or not the robot is in its HOME position  / In Home Position *)
	bErrToPlc						:BOOL;						(* $OUT[35] - Error output to PLC / Steuerungs- oder Technologiefehler aufgetreten *)
	bIOActConf						:BOOL;						(* $OUT[140] - This output is TRUE if Automatic External mode is selected and the input $I_O_ACT is TRUE. / *)
	bInWorkArea 						:BOOL;						(* $OUT[36] - Robot in work area / Roboter in Bearbeitunsbereich*)

	bForceToBase					:BOOL;						(* $OUT[10] - Move force to base position *)
	bForceToWork					:BOOL;						(* $OUT[11] - Move force to work position *)
	bCutoffToBase					:BOOL;						(* $OUT[12] - Move cutoff to base position *)
	bCutoffToWork					:BOOL;						(* $OUT[13] - Move cutoffe to work position *)

	bMEStartHeat					:BOOL;						(* $OUT[18] - Start heat *)
	bMEStopHeat					:BOOL;						(* $OUT[19] - Stop heat *)
	bMEStartExtruding					:BOOL;						(* $OUT[20] - Start extruding *)
	bMEStopExtruding					:BOOL;						(* $OUT[21] - Stop extruding *)
	bMEStartFlush 					:BOOL;						(* $OUT[22] - Start flush *)
	bMEStopFlush 					:BOOL;						(* $OUT[23] - Stop flush *)
	nMEExtrudingSpeed				:INT;						(* $OUT[100] - Extruding speed [%] *)

END_STRUCT
END_TYPE

// ---- Data types/Objects/Robot/KUKA/ST_KUKA_REF.TcDUT
TYPE ST_KUKA_REF : FB_KUKA_REF;
END_TYPE

// ---- Data types/Objects/Robot/KUKA/ST_PLCTOKUKA.TcDUT
TYPE ST_PLCTOKUKA :
STRUCT
	bDrivesOn						:BOOL;						(* $IN[140] - Switch on the robot drives / Einschalten der Roboterantriebe *)
	bDrivesOff						:BOOL;						(* $IN[141] - If this input is FALSE, Switch off the robot drives / Abschalten der Roboterantriebe *)
	bConfMess						:BOOL;						(* $IN[142] - Acknowledge error / Quittieren von Fehlermeldungen durch den Leitrechner *)
	bMoveEnable					:BOOL;						(* $IN[143] - Check the robot drives. TRUE Jogging and program execution are possible / Kontrolle der Roboterantriebe *)
	bCheckMovena					:BOOL;						(* TRUE MOVE_ENABLE monitoring is activated / Überwachung für MOVE_ENABLE *)
	bExtStart							:BOOL;						(* $IN[145] - If the I/O interface is active, this input can be set to start or continue a program / Extern Start *)
	bIOAct							:BOOL;						(* $IN[1025] - If this input is TRUE, the Automatic External interface is active. Default setting:$IN[1025]. *)
	nPgNo							:INT;						(* $IN[33] - Program number / Programmnummer *)
																(* $IN[33]  + 8 = $IN[41], PGNO_LENGTH = 8 (max. 16) *)
	bPgNoParity						:BOOL;						(* $IN[41] - Input to which the parity bit is transferred from the higher-level controller / Übertragen des Paritätsbit vom Leitrechner *)
	bPgNoValid						:BOOL;						(* $IN[42] - Input to which the command to read the program number is transferred from the higher-level controller / Einlesen der Programmnumer vom Leitrechener *)
	nOverride						:INT;						(* $IN[100] - Override *)

	bPgReset						:BOOL;						(* $IN[148] - Cancel a program / Programm abbrechen *)

	bForceInBase					:BOOL;						(* $IN[10] - Force in base position *)
	bForceInWork					:BOOL;						(* $IN[11] - Force in work position *)
	bCutoffInBase						:BOOL;						(* $IN[12] - Cutoff in base position *)
	bCutoffInWork						:BOOL;						(* $IN[13] - Cutoff in work position *)

	bMEHeat						:BOOL;						(* $IN[18] - Heat status ON = TRUE, OFF = FALSE *)
	bMEHeating						:BOOL;						(* $IN[19] - Heating status ON = TRUE, OFF = FALSE *)
	bMEHeated						:BOOL;						(* $IN[20] - Heated status ON = TRUE, OFF = FALSE *)
	bMEExtruding						:BOOL;						(* $IN[21] - Extruder status ON = TRUE, OFF = FALSE *)

	nCutOffDist						:INT;						(* $IN[50] - Distance of cutoff *)
	nExtruderOffDist					:INT;						(* $IN[66] - Distance aftre extruder is off *)
	unExtruderStartTime				:UINT;						(* $IN[82] - Extruder start time *)

END_STRUCT
END_TYPE

// ---- Data types/Objects/Robot/ST_PLCTOROBOT.TcDUT
TYPE ST_PLCTOROBOT :
STRUCT
	arbyOutput				:ARRAY[0..63] OF BYTE;
END_STRUCT
END_TYPE

// ---- Data types/Objects/Robot/ST_ROBOTTOPLC.TcDUT
TYPE ST_ROBOTTOPLC :
STRUCT
	arbyInput				:ARRAY[0..63] OF BYTE;
END_STRUCT
END_TYPE

// ---- Data types/Objects/Robot/YASKAWA/ET_YaskawaStart.TcDUT
TYPE ET_YaskawaStart :
(
	ET_YaskawaStart_eWaitExecute := 0,
	ET_YaskawaStart_eCallMasterJob,
	ET_YaskawaStart_eExternalStart,
	ET_YaskawaStart_eWfPrgDone,
	ET_YaskawaStart_eInterrupted := 196,
	ET_YaskawaStart_eDone := 197,
	ET_YaskawaStart_eError := 198,
	ET_YaskawaStart_eNoExecute := 199
);
END_TYPE

// ---- Data types/Objects/Robot/YASKAWA/ST_PLCTOYASKAWA.TcDUT
TYPE ST_PLCTOYASKAWA :
STRUCT
	bExternalStart							:BOOL;					(* If the I/O interface is active, this input can be set to start or continue a program. Only the rising edge of the signal is valid *)
	bExternalServoOn						:BOOL;					(* Switch on the robot drives. When these signals are on, the servo power supply is cut off and the manipulator stops. *)
	bCallMasterJob						:BOOL;					(* These signals have the same function as the cycle select key on the playback panel. Use the signals when desiring to change cycle specifications from the outside. *)
	bAlarmReset							:BOOL;					(* This signal clears alarms or errors when there is a minor failure,system alarm, user alarm, or user error. *)
	bReducedSpeed						:BOOL;					(* Reduced speed *)
	bExternalHold						:BOOL;					(* External hold *)

	bExternalServoOffHoldStop				:BOOL;					(* External servo off hold stop. *)
	bExternalServoOffEStop				:BOOL;					(* External servo off E-Stop *)

	bMachineError						:BOOL;					(* IN  - Machine has fault. *)
	bMachineRunning						:BOOL;					(* IN  - Machine running. *)
	bInterrupt								:BOOL;					(* IN - Interrupt;. *)

	usnOverride							:USINT;					(* IN - Override *)
	nPrgNo								:INT;					(* IN  - Automatic program number  *)

	unPipeDiameter						:UINT;					(* IN - Pipe diameter. *)
	nPipeBaseHeight						:INT;					(* IN - Pipe base height. *)
	nExtruderTowardAngle					:INT;					(* IN - Extruder toward angle deg *)
	nExtruderSideAngle					:INT;					(* IN - Extruder side angle deg *)

	bWeldingInBase						:BOOL;					(* IN - Welding in base. *)
	bWeldingInWork						:BOOL;					(* IN - Welding in work. *)
	bWeldingShoeTop					:BOOL;					(* IN - Welding shoe top. *)
	bWeldingShoeBottom					:BOOL;					(* IN - Welding shoe bottom. *)
	bWeldingHeadUnlocked				:BOOL;					(* IN - Welding head unlocked. *)
	bWeldingHeadLocked					:BOOL;					(* IN - Welding head locked. *)
	bGripperTongsOpened				:BOOL;					(* IN - Gripper tongs opened. *)
	bGripperTongsClosed					:BOOL;					(* IN - Gripper tongs closed. *)

	bWeldingInMiddle						:BOOL;					(* IN - Welding in middle position *)

END_STRUCT
END_TYPE

// ---- Data types/Objects/Robot/YASKAWA/ST_YASKAWATOPLC.TcDUT
TYPE ST_YASKAWATOPLC :
STRUCT
	bOperatingRunning						:BOOL;					(* Operating running. *)
	bServoIsOn								:BOOL;					(* Servo is on. *)
	bTopMasterJob							:BOOL;					(* Top master job. *)
	bAlarmErrorOccured						:BOOL;					(* Alarm error occured. *)
	bReducedSpeed							:BOOL;					(* Reduced speed *)
	bRemoteModeSelected					:BOOL;					(* Remote mode selected. *)
	bPlayModeSelected						:BOOL;					(* Play mode selected. *)
	bTeachModeSelected						:BOOL;					(* Teach mode selected. *)

	bHold									:BOOL;					(* Hold. *)

	bInHome									:BOOL;					(* OUT - Robot in home position. *)
	bInHeatingStationArea						:BOOL;					(* OUT - Robot in heating station area. *)
	bInFlushStationArea						:BOOL;					(* OUT - Robot in flush station area. *)
	bInLeftStationArea							:BOOL;					(* OUT - Robot in left station area. *)
	bInRightStationArea						:BOOL;					(* OUT - Robot in right station area. *)

	bPrgDone								:BOOL;					(* OUT - Program done. *)
	bPrgError								:BOOL;					(* OUT - Program done. *)
	bNotMoving								:BOOL;					(* OUT - Robot running. *)
	bNotInCrashAreaMachine					:BOOL;					(* OUT - Robot not in crash area with machine. *)

	bWeldingToBase							:BOOL;					(* OUT - Welding to base. *)
	bWeldingToWork							:BOOL;					(* OUT - Welding to work.*)
	bWeldingShoeUp							:BOOL;					(* OUT - Welding shoe move up. *)
	bWeldingShoeDown						:BOOL;					(* OUT - Welding shoe move down.*)
	bWeldingHeadUnlock						:BOOL;					(* OUT - Welding head unlock. *)
	bWeldingHeadLock						:BOOL;					(* OUT - Welding head lock. *)
	bGripperTongsOpen						:BOOL;					(* OUT - Gripper tongs open. *)
	bGripperTongsClose						:BOOL;					(* OUT - Gripper tongs close. *)

	unTargetForce							:UINT;					(* OUT - Target force [N] *)

END_STRUCT
END_TYPE

// ---- Data types/Objects/Robot/YASKAWA/ST_YASKAWA_REF.TcDUT
TYPE ST_YASKAWA_REF : FB_YASKAWA_REF;
END_TYPE

// ---- Data types/Objects/Spindle/ET_SpindleClutchStatus.TcDUT
(* Status of spindle *)

TYPE ET_SpindleClutchStatus :
(
	ET_SpindleClutchStatus_ClosedWithoutTool := 0,				(* Clutch is closed without tool *)
	ET_SpindleClutchStatus_ClosedWithTool := 1,					(* Clutch is closed with tool *)
	ET_SpindleClutchStatus_Opened := 2,						(* Clutch is opened *)
	ET_SpindleClutchStatus_RotatingNoClosed := 3,				(* Clutch rotating and not closed *)
	ET_SpindleClutchStatus_NoDefined := 999
);
END_TYPE

// ---- Data types/Objects/Spindle/PDS/ST_SpindlePDSXLA170ClutchStatus.TcDUT
TYPE ST_SpindlePDSXLA170ClutchStatus :
STRUCT
	bRotatingS1					:BOOL;						(* Spindle rotating S1 *)
	bToolNotClampedS2			:BOOL;						(* Tool not clamped S2 *)
	bToolPresentS3				:BOOL;						(* Tool present S3 *)
	bClutchInBaseS4				:BOOL;						(* Clutch in base position S4 *)
END_STRUCT
END_TYPE

// ---- Data types/Objects/Spindle/PDS/ST_SpindlePDSXLHClutchStatus.TcDUT
TYPE ST_SpindlePDSXLHClutchStatus :
STRUCT
	bToolClampedS1					:BOOL;			(* Tool clamped S1 *)
	bToolEjectedS2					:BOOL;			(* Tool present S2 *)
	bSpindleStandstillS3				:BOOL;			(* Spindle standstill S3 *)
END_STRUCT
END_TYPE

// ---- Data types/Objects/Terminal/ST_TerminalState.TcDUT
TYPE ST_TerminalState :
STRUCT
	stAdsAddr 					:ST_AmsAddr;				(* AMS Address for CoE Com *)
	bWcState					:BOOL;						(* WcState (Working Counter) *)
	unInfoState 					:UINT;						(* Info Data --> State *)
END_STRUCT
END_TYPE

// ---- Data types/Objects/TouchProbe/Renishaw/ST_TouchProbeRenishawCtrl.TcDUT
TYPE ST_TouchProbeRenishawCtrl :
STRUCT
	bMachineStartInputP1				:BOOL;			(* Machine start input [P1] *)
	bMachineStartInputP2				:BOOL;			(* Machine start input [P2] *)
	bMachineStartInputP3				:BOOL;			(* Machine start input [P3] *)
	bMachineStartInputP4				:BOOL;			(* Machine start input [P4] *)
END_STRUCT
END_TYPE

// ---- Data types/Objects/TouchProbe/Renishaw/ST_TouchProbeRenishawStatus.TcDUT
TYPE ST_TouchProbeRenishawStatus :
STRUCT
	bProbeStatus1					:BOOL;			(* Probe status 1 *)
	bLowBattery						:BOOL;			(* Low battery  *)
	bError							:BOOL;			(* Error  *)
END_STRUCT
END_TYPE

// ---- Data types/Objects/VFD/ST_PLCTOVFD.TcDUT
TYPE ST_PLCTOVFD :
STRUCT
	bEnable							:BOOL;			(* Enable controller *)
	bFaultReset						:BOOL;			(* Acknowledgment for faults of the device state machine. *)
	bForwardStop					:BOOL;			(* Counterclockwise rotation moving. *)
	bReverseStop					:BOOL;			(* Clockwise rotation moving. *)
	bJog							:BOOL;			(* Jog command. *)
	bExtError							:BOOL;			(* External error signal. *)
	nSetMotorSpeed					:INT;			(* Relative speed reference value *)
	bReserve1						:BOOL;			(* Reserve 1. *)
	bReserve2						:BOOL;			(* Reserve 2. *)
END_STRUCT
END_TYPE

// ---- Data types/Objects/VFD/ST_VFDTOPLC.TcDUT
TYPE ST_VFDTOPLC :
STRUCT
	bEnabled						:BOOL;			(* The drive is on. *)
	bOperational						:BOOL;			(* The drive is ready for operation. *)
	bBrakeError						:BOOL;			(* Brake device error *)
	bDummy							:BOOL;
	nCurrentMotorSpeed				:INT;			(* Current motor speed *)
END_STRUCT
END_TYPE

// ---- Data types/Objects/VFD/ST_VFD_AXIS_REF.TcDUT
TYPE ST_VFD_AXIS_REF : FB_VFD_Axis_REF;
END_TYPE

// ---- Data types/Objects/VFD/ST_VFD_DRIVE_REF.TcDUT
TYPE ST_VFD_DRIVE_REF : FB_VFD_Drive_REF;
END_TYPE

// ---- POUs/Tc3 Objects/Alarm/ET_AlarmType_1.TcDUT
{attribute 'qualified_only'}
{attribute 'strict'}
TYPE ET_AlarmType_1 : 
(
	eIdle := 0,
	eFatalError := 1,
	eError := 2,
	eWarning := 3,
	eMessage := 4,
	eHint := 5	
)INT;
END_TYPE

// ---- POUs/Tc3 Objects/Alarm/ST_AlarmIn_1.TcDUT
TYPE ST_AlarmIn_1 :
STRUCT
	arbFatalError		:ARRAY[0..nALARM_MAX_NO] OF ST_AlarmProperties;
	arbError			:ARRAY[0..nALARM_MAX_NO] OF ST_AlarmProperties;
	arbWarning			:ARRAY[0..nALARM_MAX_NO] OF ST_AlarmProperties;
	arbMessage			:ARRAY[0..nALARM_MAX_NO] OF ST_AlarmProperties;
	arbHint				:ARRAY[0..nALARM_MAX_NO] OF ST_AlarmProperties;
END_STRUCT
END_TYPE

// ---- POUs/Tc3 Objects/Alarm/ST_AlarmOut_1.TcDUT
TYPE ST_AlarmOut_1 :
STRUCT
	arbFatalError		:ARRAY[0..nALARM_MAX_NO] OF ST_AlarmProperties;
	arbError			:ARRAY[0..nALARM_MAX_NO] OF ST_AlarmProperties;
	arbWarning			:ARRAY[0..nALARM_MAX_NO] OF ST_AlarmProperties;
	arbMessage			:ARRAY[0..nALARM_MAX_NO] OF ST_AlarmProperties;
	arbHint				:ARRAY[0..nALARM_MAX_NO] OF ST_AlarmProperties;
	bFatalError			:BOOL;				(* Fatal error in group / Fataler Fehler in der Gruppe *)
	bError				:BOOL;				(* Error in group / Fehler in der Gruppe *)
	bWarning			:BOOL;				(* Warning in group / Warnung  in der Gruppe *)
	bMessage			:BOOL;				(* Message in group / Meldung in der Gruppe *)
	bHint				:BOOL;				(* Hint in group / Hint in der Gruppe *)
END_STRUCT
END_TYPE

// ---- POUs/Tc3 Objects/Alarm/ST_AlarmProperties_1.TcDUT
TYPE ST_AlarmProperties_1 :
STRUCT
	bActive				:BOOL;				(* Alarm on *)
	{attribute 'hide'} 
	dtDateTime			:DATE_AND_TIME ;	(* Alarm time stamp *)
	{attribute 'hide'} 
	enType				:ET_AlarmType;		(* Alarm type *)
	dnCode				:DINT;				(* Alarm code *)
END_STRUCT
END_TYPE

// ---- POUs/Tc3 Objects/Alarm/ST_AlarmRef_1.TcDUT
TYPE ST_AlarmRef_1 :
STRUCT
	stControl				:ST_AlarmOut;
	stManual				:ST_AlarmOut;
	//stMaintenance			:ST_AlarmOut;
	stHome					:ST_AlarmOut;
	stAuto					:ST_AlarmOut;
END_STRUCT
END_TYPE

// ---- POUs/Tc3 Objects/Alarm/ST_Alarm_1.TcDUT
TYPE ST_Alarm_1 :
STRUCT
	bFatalError			:BOOL;				(* Fatal error in group / Fataler Fehler in der Gruppe *)
	bError				:BOOL;				(* Error in group / Fehler in der Gruppe *)
	bWarning			:BOOL;				(* Warning in group / Warnung  in der Gruppe *)
	bMessage			:BOOL;				(* Message in group / Meldung in der Gruppe *)
	bHint				:BOOL;				(* Hint in group / Hint in der Gruppe *)
END_STRUCT
END_TYPE

// ---- POUs/Tc3 Objects/Automation/OperationMode/ET_MachineMode_1.TcDUT
(* Machine operating mode *)
TYPE ET_MachineMode_1 :
(
	ET_MachineMode_eUndefined := 0,
	ET_MachineMode_eAutomatic := 1,
	ET_MachineMode_eCycle := 2,
	ET_MachineMode_eStepping := 3,
	ET_MachineMode_eHome := 4,
	ET_MachineMode_eManual := 5,
	ET_MachineMode_eMaintenance := 6,
	ET_MachineMode_eDryRun := 7,
	ET_MachineMode_eMDI := 8,
	ET_MachineMode_eIdle := 10
);
END_TYPE

// ---- POUs/Tc3 Objects/Automation/OperationMode/ET_MachineState_1.TcDUT
(* Machine state *)
TYPE ET_MachineState_1 :
(
	ET_MachineState_eUndefined := 0,
	ET_MachineState_eAutoExe := 1,
	ET_MachineState_eAutoSteppingExe := 2,
	ET_MachineState_eAutoSteppingNoExe := 3,
	ET_MachineState_eHomeExe := 4,
	ET_MachineState_eHomeRefExe := 5,
	ET_MachineState_eMaintenanceExe := 6,
	ET_MachineState_eIdle := 10
) ;
END_TYPE

// ---- POUs/Tc3 Objects/Automation/OperationMode/ET_MaintenanceType.TcDUT
(* Machine operating mode *)
TYPE ET_MaintenanceType :
(
	ET_MaintenanceType_eUndefined := 0,
	ET_MaintenanceType_eCooling := 1,
	ET_MaintenanceType_eCGK := 2
);
END_TYPE

// ---- POUs/Tc3 Objects/Communication/TCPIP/ET_TCPIP_ConnectionState.TcDUT
TYPE ET_TCPIP_ConnectionState :
(
	ET_TCPIP_ConnState_eIdle := 0,
	ET_TCPIP_ConnState_eConnect,
	ET_TCPIP_ConnState_eDataExchsnge,
	ET_TCPIP_ConnState_eDisconnect
);
END_TYPE

// ---- POUs/Tc3 Objects/Diagnostic/Terminal/ST_TerminalState_1.TcDUT
TYPE ST_TerminalState_1 :
STRUCT
	stAdsAddr 					:ST_AmsAddr;				(* AMS Address for CoE Com *)
	bWcState					:BOOL;						(* WcState (Working Counter) *)
	unInfoState 					:UINT;						(* Info Data --> State *)
END_STRUCT
END_TYPE

// ---- POUs/Tc3 Objects/Engineering/External set value generator/ET_ExtSetpoint.TcDUT
TYPE ET_ExtSetpoint :
(
	ET_ExtSetpoint_eWaitExecute := 0,
	ET_ExtSetpoint_eEnableExtSetPointGenerator := 5,
	ET_ExtSetpoint_eDisableExtSetPointGenerator := 10,
	ET_ExtSetpoint_eDone := 197,
	ET_ExtSetpoint_eError := 198,
	ET_ExtSetpoint_eNoExecute := 199
);
END_TYPE

// ---- POUs/Tc3 Objects/ExternalHardware/Gefran/ET_GFX4IR_1.TcDUT
TYPE ET_GFX4IR_1 :
(
	ET_GFX4IRState_eWaitExecute := 0,
	ET_GFX4IRState_eCtrlOn,
	ET_GFX4IRState_eCtrlOff,
	ET_GFX4IRState_eDone := 197,
	ET_GFX4IRState_eError := 198,
	ET_GFX4IRState_eNoExecute := 199
);
END_TYPE

// ---- POUs/Tc3 Objects/ExternalHardware/Gefran/ST_GFX4IRTOPLC_1.TcDUT
(* Communikation structure from plc to gefran *)

TYPE ST_GFX4IRTOPLC_1 :
STRUCT
	nProcessVariable			:INT;
	wControllerStatus			:WORD;
	nOutputPower				:INT;
	wAmmeterInputOn				:WORD;
END_STRUCT
END_TYPE

// ---- POUs/Tc3 Objects/ExternalHardware/Gefran/ST_GFX4IR_REF_1.TcDUT
TYPE ST_GFX4IR_REF_1 : FB_GFX4IR_REF;
END_TYPE

// ---- POUs/Tc3 Objects/ExternalHardware/Gefran/ST_PLCTOGFX4IR_1.TcDUT
(* Communikation structure from gefran to plc *)

TYPE ST_PLCTOGFX4IR_1 :
STRUCT
	nLocalSetPoint			:INT;
	nManualOutput			:WORD;
	wControllerStatus		:WORD;
END_STRUCT
END_TYPE

// ---- POUs/Tc3 Objects/ExternalHardware/KUKA/ET_KukaStart_1.TcDUT
TYPE ET_KukaStart_1 :
(
	ET_KukaStart_eWaitExecute := 0,
	ET_KukaStart_eExtStart,
	ET_KukaStart_eWfInHome,
	ET_KukaStart_eWfPgNoReq,
	ET_KukaStart_ePgNoParity,
	ET_KukaStart_ePgNoValid,
	ET_KukaStart_eWfProgFinish,
	ET_KukaStart_eDone := 197,
	ET_KukaStart_eError := 198,
	ET_KukaStart_eNoExecute := 199
);
END_TYPE

// ---- POUs/Tc3 Objects/ExternalHardware/KUKA/ST_KUKATOPLC_1.TcDUT
TYPE ST_KUKATOPLC_1 :
STRUCT
	bStopMess						:BOOL;						(* $OUT[1010] - Any message occurring which requires the robot to be stopped / Störung Roboter *)
	bPgNoReq						:BOOL;						(* $OUT[33] - A change of signal requests the higher-level controller to send a program number / PGNO Req-Signalwechsel fordert Leitrechner Programmnr. zu senden *)
	bApplRun						:BOOL;						(* $OUT[34] - Program is currently being executed / TRUE wenn Programm abgearbeitet wird *)
	bPeriRdy						:BOOL;						(* $OUT[1012] - Robot drives are switched on / TRUE wenn Roboterantriebe eingeschaltet *)
	bAlarmStop						:BOOL;						(* $OUT[1013] - Emergency stop / Not Aus *)
	bUserSafe						:BOOL;						(* $OUT[1011] - If the safety fence monitoring switch is opened (AUT mode) or an enabling switch is released (T1 or T2 mode). / Abfrage Schutzgitter(Auto)/Zustimmungsschalter(Test) *)
	bT1								:BOOL;						(* $OUT[993] - Operating mode T1 / Betriebsart T1 *)
	bT2								:BOOL;						(* $OUT[994] - Operating mode T2/ Betriebsart T2 *)
	bAut								:BOOL;						(* $OUT[995] - Operating mode Aut / Betriebsart Aut *)
	bExt								:BOOL;						(* $OUT[996] - Operating mode Ext / Betriebsart Ext *)
	bOnPath							:BOOL;						(* $OUT[997] - Set as long as the robot stays on its programmed path / TRUE solange sich Rob. auf programmierten Bahn befindet *)
	bProAct							:BOOL;						(* $OUT[1021] - Whenever a process is active / Programmbearbeitung aktiv *)
	bInHome							:BOOL;						(* $OUT[1000] - Whether or not the robot is in its HOME position  / In Home Position *)
	arbInHome						:ARRAY[1..5] OF BOOL;		(* $OUT[1003..1007] - Whether or not the robot is in its HOME position  / In Home Position *)
	bErrToPlc						:BOOL;						(* $OUT[35] - Error output to PLC / Steuerungs- oder Technologiefehler aufgetreten *)
	bIOActConf						:BOOL;						(* $OUT[140] - This output is TRUE if Automatic External mode is selected and the input $I_O_ACT is TRUE. / *)
	bInWorkArea 						:BOOL;						(* $OUT[36] - Robot in work area / Roboter in Bearbeitunsbereich*)

	bForceToBase					:BOOL;						(* $OUT[10] - Move force to base position *)
	bForceToWork					:BOOL;						(* $OUT[11] - Move force to work position *)
	bCutoffToBase					:BOOL;						(* $OUT[12] - Move cutoff to base position *)
	bCutoffToWork					:BOOL;						(* $OUT[13] - Move cutoffe to work position *)

	bMEStartHeat					:BOOL;						(* $OUT[18] - Start heat *)
	bMEStopHeat					:BOOL;						(* $OUT[19] - Stop heat *)
	bMEStartExtruding					:BOOL;						(* $OUT[20] - Start extruding *)
	bMEStopExtruding					:BOOL;						(* $OUT[21] - Stop extruding *)
	bMEStartFlush 					:BOOL;						(* $OUT[22] - Start flush *)
	bMEStopFlush 					:BOOL;						(* $OUT[23] - Stop flush *)
	nMEExtrudingSpeed				:INT;						(* $OUT[100] - Extruding speed [%] *)

END_STRUCT
END_TYPE

// ---- POUs/Tc3 Objects/ExternalHardware/KUKA/ST_KUKA_REF_1.TcDUT
TYPE ST_KUKA_REF_1 : FB_KUKA_REF;
END_TYPE

// ---- POUs/Tc3 Objects/ExternalHardware/KUKA/ST_PLCTOKUKA_1.TcDUT
TYPE ST_PLCTOKUKA_1 :
STRUCT
	bDrivesOn						:BOOL;						(* $IN[140] - Switch on the robot drives / Einschalten der Roboterantriebe *)
	bDrivesOff						:BOOL;						(* $IN[141] - If this input is FALSE, Switch off the robot drives / Abschalten der Roboterantriebe *)
	bConfMess						:BOOL;						(* $IN[142] - Acknowledge error / Quittieren von Fehlermeldungen durch den Leitrechner *)
	bMoveEnable					:BOOL;						(* $IN[143] - Check the robot drives. TRUE Jogging and program execution are possible / Kontrolle der Roboterantriebe *)
	bCheckMovena					:BOOL;						(* TRUE MOVE_ENABLE monitoring is activated / Überwachung für MOVE_ENABLE *)
	bExtStart							:BOOL;						(* $IN[145] - If the I/O interface is active, this input can be set to start or continue a program / Extern Start *)
	bIOAct							:BOOL;						(* $IN[1025] - If this input is TRUE, the Automatic External interface is active. Default setting:$IN[1025]. *)
	nPgNo							:INT;						(* $IN[33] - Program number / Programmnummer *)
																(* $IN[33]  + 8 = $IN[41], PGNO_LENGTH = 8 (max. 16) *)
	bPgNoParity						:BOOL;						(* $IN[41] - Input to which the parity bit is transferred from the higher-level controller / Übertragen des Paritätsbit vom Leitrechner *)
	bPgNoValid						:BOOL;						(* $IN[42] - Input to which the command to read the program number is transferred from the higher-level controller / Einlesen der Programmnumer vom Leitrechener *)
	nOverride						:INT;						(* $IN[100] - Override *)

	bPgReset						:BOOL;						(* $IN[148] - Cancel a program / Programm abbrechen *)

	bForceInBase					:BOOL;						(* $IN[10] - Force in base position *)
	bForceInWork					:BOOL;						(* $IN[11] - Force in work position *)
	bCutoffInBase						:BOOL;						(* $IN[12] - Cutoff in base position *)
	bCutoffInWork						:BOOL;						(* $IN[13] - Cutoff in work position *)

	bMEHeat						:BOOL;						(* $IN[18] - Heat status ON = TRUE, OFF = FALSE *)
	bMEHeating						:BOOL;						(* $IN[19] - Heating status ON = TRUE, OFF = FALSE *)
	bMEHeated						:BOOL;						(* $IN[20] - Heated status ON = TRUE, OFF = FALSE *)
	bMEExtruding						:BOOL;						(* $IN[21] - Extruder status ON = TRUE, OFF = FALSE *)

	nCutOffDist						:INT;						(* $IN[50] - Distance of cutoff *)
	nExtruderOffDist					:INT;						(* $IN[66] - Distance aftre extruder is off *)
	unExtruderStartTime				:UINT;						(* $IN[82] - Extruder start time *)

END_STRUCT
END_TYPE

// ---- POUs/Tc3 Objects/ExternalHardware/Periphery/ST_PERIPHERY_REF_1.TcDUT
TYPE ST_PERIPHERY_REF_1 : FB_PERIPHERY_REF;
END_TYPE

// ---- POUs/Tc3 Objects/ExternalHardware/Periphery/ST_PLC01TOPLC02.TcDUT
TYPE ST_PLC01TOPLC02 :
STRUCT
	etMachineMode						:ET_MachineMode;			(* Machine mode *)
	etMachineState						:ET_MachineState;			(* Machine state *)
	etMaintenanceType					:ET_MaintenanceType;		(* Maintenance type *)
	bModeAutomatic						:BOOL;						(* Machine mode automatic *)
	bModeHome							:BOOL;						(* Machine mode home *)
	bModeMaintenance					:BOOL;						(* Machine mode maintenance *)
	bModeManual							:BOOL;						(* Machine mode manual *)
	bMachineRunning						:BOOL;						(* Machine running / Maschine lauft *)
	bMachineStandstill					:BOOL;						(* Machine standstill / Maschin steht *)
	bMachinePurge						:BOOL;						(* Machine purge *)
	bConfirmAlarm						:BOOL;						(* Confirm alarm *)
	rOverride							:REAL;						(* Override *)

END_STRUCT
END_TYPE

// ---- POUs/Tc3 Objects/ExternalHardware/Periphery/ST_PLC02TOPLC01.TcDUT
TYPE ST_PLC02TOPLC01 :
STRUCT
	bSafetyCompleted					:BOOL;				(* Safety completed *)
	bManualCompleted					:BOOL;				(* Manual completed *)
	bHomeCompleted						:BOOL;				(* Home completed / Grundsrellung ausgeführt *)
	bAutoCompleted						:BOOL;				(* Automatic completed / Automatik beendet *)
	bMaintenanceCompleted				:BOOL;				(* Maintenance completed / Maintenance beendet*)
	bFatalError							:BOOL;				(* Fatal error in group / Fataler Fehler in der Gruppe *)
	bError								:BOOL;				(* Error in group / Fehler in der Gruppe *)
	bWarning							:BOOL;				(* Warning in group / Warnung  in der Gruppe *)
	bMessage							:BOOL;				(* Message in group / Meldung in der Gruppe *)
	bHint								:BOOL;				(* Hint in group / Hint in der Gruppe *)
	bAllDoorsClosed						:BOOL;				(* All doors closed / Alle Türen geschlossen *)
	bAllDoorsClosedLocked				:BOOL;				(* All doors closed and locked / Alle Türen geschlossen und verrrigelt *)
	
	bHazard								:BOOL;				(* Hazard *)
END_STRUCT
END_TYPE

// ---- POUs/Tc3 Objects/ExternalHardware/Periphery/ST_PLC02TOPLC03.TcDUT
TYPE ST_PLC02TOPLC03 :
STRUCT	
	bShuttleWeldingReq					:BOOL;						(* Shuttle request *)
	bShuttleMillingAck					:BOOL;						(* Shuttle acknowledge *)
	lrShuttleMillingActPos				:LREAL;						(* Actual position of shuttel [mm] *)
	lrShuttleMillingSetPos				:LREAL;						(* Set position of shuttel [mm] *)
	
	arbMillingActive					:ARRAY[0..GVL_FB_LoadFromFile.usnFileArrayMaxDimR] OF BOOL; 			(* Process milling active *)	
	arbMillingDone						:ARRAY[0..GVL_FB_LoadFromFile.usnFileArrayMaxDimR] OF BOOL; 			(* Process milling done *)	
	
	bMillingDriveEnabled				:BOOL;						(* Drive enabled *)
	bMillingDriveEnable					:BOOL;						(* Drive enable *)
END_STRUCT
END_TYPE

// ---- POUs/Tc3 Objects/ExternalHardware/Periphery/ST_PLC03TOPLC02.TcDUT
TYPE ST_PLC03TOPLC02 :
STRUCT
	bShuttleMillingReq					:BOOL;						(* Shuttle request *)
	bShuttleWeldingAck					:BOOL;						(* Shuttle acknowledge *)
	lrShuttleWeldingActPos				:LREAL;						(* Actual position of shuttel [mm] *)
	lrShuttleWeldingSetPos				:LREAL;						(* Set position of shuttel [mm] *)
	
	arbWeldingActive					:ARRAY[0..GVL_FB_LoadFromFile.usnFileArrayMaxDimR] OF BOOL; 			(* Process welding active *)	
	arbWeldingDone						:ARRAY[0..GVL_FB_LoadFromFile.usnFileArrayMaxDimR] OF BOOL; 			(* Process welding done *)	
	
	bWeldingDriveEnabled				:BOOL;						(* Drive enabled *)
	bWeldingDriveEnable					:BOOL;						(* Drive enable *)
	
END_STRUCT
END_TYPE

// ---- POUs/Tc3 Objects/ExternalHardware/Robot/ST_PLCTOROBOT_1.TcDUT
TYPE ST_PLCTOROBOT_1 :
STRUCT
	arbyOutput				:ARRAY[0..31] OF BYTE;
END_STRUCT
END_TYPE

// ---- POUs/Tc3 Objects/ExternalHardware/Robot/ST_ROBOTTOPLC_1.TcDUT
TYPE ST_ROBOTTOPLC_1 :
STRUCT
	arbyInput				:ARRAY[0..31] OF BYTE;
END_STRUCT
END_TYPE

// ---- POUs/Tc3 Objects/ExternalHardware/YASKAWA/ET_YaskawaStart_1.TcDUT
TYPE ET_YaskawaStart_1 :
(
	ET_YaskawaStart_eWaitExecute := 0,
	ET_YaskawaStart_eCallMasterJob,
	ET_YaskawaStart_eExternalStart,
	ET_YaskawaStart_eWfPrgDone,
	ET_YaskawaStart_eDone := 197,
	ET_YaskawaStart_eError := 198,
	ET_YaskawaStart_eNoExecute := 199
);
END_TYPE

// ---- POUs/Tc3 Objects/ExternalHardware/YASKAWA/ST_PLCTOYASKAWA_1.TcDUT
TYPE ST_PLCTOYASKAWA_1 :
STRUCT
	bExternalStart							:BOOL;					(* If the I/O interface is active, this input can be set to start or continue a program. Only the rising edge of the signal is valid *)
	bExternalServoOn						:BOOL;					(* Switch on the robot drives. When these signals are on, the servo power supply is cut off and the manipulator stops. *)
	bCallMasterJob						:BOOL;					(* These signals have the same function as the cycle select key on the playback panel. Use the signals when desiring to change cycle specifications from the outside. *)
	bAlarmReset							:BOOL;					(* This signal clears alarms or errors when there is a minor failure,system alarm, user alarm, or user error. *)
	bReducedSpeed						:BOOL;					(* Reduced speed *)
	bExternalHold						:BOOL;					(* External hold *)

	bExternalServoOffHoldStop				:BOOL;					(* External servo off hold stop. *)
	bExternalServoOffEStop				:BOOL;					(* External servo off E-Stop *)

	nOverride							:INT;					(* Override *)

	bMachineError						:BOOL;					(* IN  - Machine has fault. *)
	bMachineRunning						:BOOL;					(* IN  - Machine running. *)
	bAxisClampingPosA					:BOOL;					(* IN  - Axis clamping in positon A. *)
	bAxisClampingPosB					:BOOL;					(* IN  - Axis clamping in positon B. *)

	bSpindlePresent						:BOOL;					(* IN  - Spindle present. *)
	bFurrowingPresent					:BOOL;					(* IN  - Furrowing present. *)

	bHeadSocketAirOpened				:BOOL;					(* IN  - Head socket air opened. *)
	bHeadSocketAirClosed				:BOOL;					(* IN  - Head socket air closed. *)
	bHeadUnDocked						:BOOL;					(* IN  - Head undocked. *)
	bHeadDocked						:BOOL;					(* IN  - Head docked. *)
	bGetHeadNestDone					:BOOL;					(* IN  - Get head nest done. *)

	bToolStorageHoodOpened				:BOOL;					(* IN  - Tool storage hood opened. *)
	bToolStorageHoodClosed				:BOOL;					(* IN  - Tool storage hood closed. *)
	bGetToolNestDone					:BOOL;					(* IN  - Get tool nest done. *)

	bSpindleBitClutchOpened				:BOOL;					(* IN  - Spindle bit clutch opened. *)
	bSpindleBitClutchClosed				:BOOL;					(* IN  - Spindle bit clutch closed. *)
	bSpindleBitClutchClosedWithTool		:BOOL;					(* IN  - Spindle bit clutch with tool closed. *)
	bSpindleNotMoving					:BOOL;					(* IN  - Spindle not moving. *)
	bSpindleReady						:BOOL;					(* IN  - Spindle ready. *)
	bSpindlePurgeOpened					:BOOL;					(* IN -  Spindle purge opened. *)
	bSpindlePurgeClosed					:BOOL;					(* IN -  Spindle purge closed. *)

	bFurrowingHeadUnlocked				:BOOL;					(* IN  - Furrowing head unlocked. *)
	bFurrowingHeadLocked				:BOOL;					(* IN  - Furrowing head locked. *)
	bFurrowingHeadCutterOpened			:BOOL;					(* IN  - Furrowing head cutter opened. *)
	bFurrowingHeadCutterClosed			:BOOL;					(* IN  - Furrowing head cutter closed. *)

	bPipeMeasurementEn					:BOOL;					(* IN - Enable pipe measurement. *)
	bTouchProbeStatus1					:BOOL;					(* IN  - Touch probe status 1. *)

	unToolNestAct						:UINT;					(* IN  - Current tool nest number *)
	unToolNestPrv						:UINT;					(* IN  - Previous tool nest number *)
	unHeadNestAct						:UINT;					(* IN  - Current head nest number *)
	unHeadNestPrv						:UINT;					(* IN  - Previous head nest number *)

	nPrgNo								:INT;					(* IN  - Automatic program number  *)

	unPipeDiameter						:UINT;					(* IN - Pipe diameter *)
	unPipeLengthA						:UINT;					(* IN - Pipe length A *)
	unPipeLengthB						:UINT;					(* IN - Pipe length B *)

	unOverride							:UINT;					(* IN - Override *)
END_STRUCT
END_TYPE

// ---- POUs/Tc3 Objects/ExternalHardware/YASKAWA/ST_YASKAWATOPLC_1.TcDUT
TYPE ST_YASKAWATOPLC_1 :
STRUCT
	bOperatingRunning						:BOOL;					(* Operating running. *)
	bServoIsOn								:BOOL;					(* Servo is on. *)
	bTopMasterJob							:BOOL;					(* Top master job. *)
	bAlarmErrorOccured						:BOOL;					(* Alarm error occured. *)
	bReducedSpeed							:BOOL;					(* Reduced speed *)
	bRemoteModeSelected					:BOOL;					(* Remote mode selected. *)
	bPlayModeSelected						:BOOL;					(* Play mode selected. *)
	bTeachModeSelected						:BOOL;					(* Teach mode selected. *)

	bHold									:BOOL;					(* Hold. *)

	bInHome									:BOOL;					(* OUT - Robot in home position. *)
	bPrgDone								:BOOL;					(* OUT - Program done. *)
	bNotInCrashAreaMachine					:BOOL;					(* OUT - Robot not in crash area with machine. *)
	bNotMoving								:BOOL;					(* OUT - Robot running. *)

	bHeadSocketAirOpen						:BOOL;					(* OUT - Head socket air open. *)
	bHeadSocketAirClose						:BOOL;					(* OUT - Head socket air close.*)
	bHeadUnDock							:BOOL;					(* OUT - Head undock. *)
	bHeadDock								:BOOL;					(* OUT - Head dock.*)
	bExeHeadNest							:BOOL;					(* OUT - Execute head nest . *)

	bToolStorageHoodOpen					:BOOL;					(* OUT - Tool storage hood open. *)
	bToolStorageHoodClose					:BOOL;					(* OUT - Tool storage hood close. *)
	bExeToolNest							:BOOL;					(* OUT - Execute tool nest . *)

	bSpindleBitClutchOpen						:BOOL;					(* OUT - Spindle bit clutch open. *)
	bSpindleBitClutchClose					:BOOL;					(* OUT - Spindle bit clutch close.*)
	bSpindleStart								:BOOL;					(* OUT - Spindle start. *)
	bSpindleStop								:BOOL;					(* OUT - Spindle stop. *)
	bSpindlePurgeOpen						:BOOL;					(* OUT - Spindle purge open *)
	bSpindlePurgeClose						:BOOL;					(* OUT - Spindle purge close *)

	bFurrowingHeadUnlock					:BOOL;					(* OUT - Furrowing head unlock. *)
	bFurrowingHeadLock						:BOOL;					(* OUT - Furrowing head lock.*)
	bFurrowingHeadCutterOpen					:BOOL;					(* OUT - Furrowing head cutter open. *)
	bFurrowingHeadCutterClose				:BOOL;					(* OUT - Furrowing head cutter close.*)

	bStartTouchProbeP1						:BOOL;					(* OUT - Start touch probe P1. *)

	unHeadNo								:UINT;					(* OUT - Head number. *)
	unToolNo								:UINT;					(* OUT - Hool number. *)
	nSpindleSpeed							:INT;					(* OUT - Spindle speed. *)

END_STRUCT
END_TYPE

// ---- POUs/Tc3 Objects/ExternalHardware/YASKAWA/ST_YASKAWA_REF_1.TcDUT
TYPE ST_YASKAWA_REF_1 : FB_YASKAWA_REF;
END_TYPE

// ---- POUs/Tc3 Objects/File/CSV/ET_CSV_State.TcDUT
TYPE ET_CSV_State :
(
	ET_CSV_State_eWaitExecute := 0,
	ET_CSV_State_eCreateDir,
	ET_CSV_State_eChkCreateDir,
	ET_CSV_State_eFileOpen,
	ET_CSV_State_eChkFileOpen,
	ET_CSV_State_eConvertRecord,
	ET_CSV_State_eFilePuts,
	ET_CSV_State_eChkFilePuts,
	ET_CSV_State_eFileGets,
	ET_CSV_State_eChkFileGets,
	ET_CSV_State_eParseSingleRecord,
	ET_CSV_State_eFileClose,
	ET_CSV_State_eChkFileClose,
	ET_CSV_State_eDone := 197,
	ET_CSV_State_eError := 198,
	ET_CSV_State_eNoExecute := 199
);
END_TYPE

// ---- POUs/Tc3 Objects/File/TXT/ET_LoadFromFile_1.TcDUT

TYPE ET_LoadFromFile_1 :
(
	ET_LoadFromFile_eWaitExecute := 0,
	ET_LoadFromFile_eFileName,
	ET_LoadFromFile_eChkFileExist,
	ET_LoadFromFile_eFileOpen,
	ET_LoadFromFile_eChkFileOpen,
	ET_LoadFromFile_eReadData,
	ET_LoadFromFile_eChkReadData,
	ET_LoadFromFile_eFileClose,
	ET_LoadFromFile_eChkFileClose,
	ET_LoadFromFile_eDone := 197,
	ET_LoadFromFile_eError := 198,
	ET_LoadFromFile_eNoExecute := 199
);
END_TYPE

// ---- POUs/Tc3 Objects/Logger/ST_LoggerVar_1.TcDUT
TYPE ST_LoggerVar_1 :
STRUCT
	udnCycleNo		:UDINT;
	sTimeStamp		:STRING(15);			(* Alarm time stamp *)
	arsLogVars		:ARRAY[1..GVL_Logger.unNUM_OF_LOG_VAR] OF STRING(10);
END_STRUCT
END_TYPE

// ---- POUs/Tc3 Objects/Logger/ST_Logger_1.TcDUT
TYPE ST_Logger_1 :
STRUCT
	arstLoggerWaitInterrupt					:ARRAY[1..GVL_Logger.unLOG_BEFOR_MAX_NO] OF ST_LoggerVar;
	arstLoggerDuringInterrupt				:ARRAY[1..GVL_Logger.unLOG_DURING_MAX_NO] OF ST_LoggerVar;
	arstLoggerAfterInterrupt					:ARRAY[1..GVL_Logger.unLOG_AFTER_MAX_NO] OF ST_LoggerVar;
END_STRUCT
END_TYPE

// ---- POUs/Tc3 Objects/Measurements/Counter/ST_TimeHoursCounter_1.TcDUT
TYPE ST_TimeHoursCounter_1 :
STRUCT
	lrAllOverHours					:LREAL; 							(* All over counter hours *)
	lrAfterResetHours					:LREAL; 							(* Counter hours since last reset *)
END_STRUCT
END_TYPE

// ---- POUs/Tc3 Objects/Measurements/ST_Time_1.TcDUT
TYPE ST_Time_1 :
STRUCT
	dwSec				:DWORD; 						(* Time in 1 [s] *)
	dwDeciSec			:DWORD; 						(* Time in deci 0.1 [s] *)
	dwCentiSec			:DWORD; 						(* Time in centi 0.01 [s] *)
	dwMiliSec			:DWORD; 						(* Time in mili 0.001 [s] *)
END_STRUCT
END_TYPE

// ---- POUs/Tc3 Objects/Safety/Fieldbus/ST_FieldbusStatus_1.TcDUT
TYPE ST_FieldbusStatus_1 :
STRUCT
	wFrmXWcState				:WORD; (* link to task related ethercat frame state FrmXWcState *)
	nMasterDeviceId				:UINT;
	nMasterSlaveCount			:UINT;
	nMasterDevState				:UINT;
	arrMasterNetId				:T_AmsNetIdArr;
	nMasterSlaveCountCfg			:UINT;
END_STRUCT
END_TYPE

// ---- POUs/Tc3 Objects/Signals/Generators/ST_Blinker_1.TcDUT
TYPE ST_Blinker_1 :
STRUCT	
	Q0					:BOOL; 						(* Divider output / 2 *)
	Q1					:BOOL; 						(* Divider output / 4 *)
	Q2					:BOOL; 						(* Divider output / 8 *)
	Q3					:BOOL; 						(* Divider output / 16 *)
	Q4					:BOOL; 						(* Divider output / 32 *)
	Q5					:BOOL; 						(* Divider output / 64 *)
	Q6					:BOOL; 						(* Divider output / 128 *)
	Q7					:BOOL; 						(* Divider output / 256 *)
END_STRUCT
END_TYPE

// ---- POUs/Tc3 Objects/Signals/Ramp Generators/ET_RampGenerator_1.TcDUT
TYPE ET_RampGenerator_1 :
(
	ET_RampGenerator_eWaitExecute := 0,
	ET_RampGenerator_eRunning := 5,
	ET_RampGenerator_eWaiting := 10,
	ET_RampGenerator_eDone := 197,
	ET_RampGenerator_eError := 198,
	ET_RampGenerator_eNotExecute := 199
);
END_TYPE

// ---- POUs/Tc3 Objects/Traceability/ET_TRACE_State.TcDUT
TYPE ET_TRACE_State :
(
	ET_TRACE_State_eWaitExecute := 0,
	ET_TRACE_State_eGetData,
	ET_TRACE_State_eDataWrite,
	ET_TRACE_State_eWfDataWrite,
	ET_TRACE_State_eDone := 197,
	ET_TRACE_State_eError := 198,
	ET_TRACE_State_eNoExecute := 199
);
END_TYPE

// ---- Global Variables/Alarms/GVL_Gr00Alarm.TcGVL
{attribute 'Tc2GvlVarNames'}
VAR_GLOBAL
	stgGr00Alarm			:ST_AlarmRef;
END_VAR

// ---- Global Variables/Alarms/GVL_Gr01Alarm.TcGVL
{attribute 'Tc2GvlVarNames'}
VAR_GLOBAL
	stgGr01Alarm			:ST_AlarmRef;
END_VAR

// ---- Global Variables/Alarms/GVL_Gr02Alarm.TcGVL
{attribute 'Tc2GvlVarNames'}
VAR_GLOBAL
	stgGr02Alarm			:ST_AlarmRef;
END_VAR

// ---- Global Variables/Alarms/GVL_Gr05Alarm.TcGVL
{attribute 'Tc2GvlVarNames'}
VAR_GLOBAL
	stgGr05Alarm			:ST_AlarmRef;
END_VAR

// ---- Global Variables/Basics/GVL_FB_CheckArrayBounds.TcGVL
{attribute 'Tc2GvlVarNames'}
VAR_GLOBAL
	(*fbCheckArrayBounds: FB_CheckArrayBounds;*)

END_VAR

// ---- Global Variables/Basics/GVL_FB_CheckDivRealInfo.TcGVL
{attribute 'Tc2GvlVarNames'}
VAR_GLOBAL
	(*fbCheckDivRealInfo: FB_CheckDivRealInfo;*)
END_VAR

// ---- Global Variables/Config/GVL_Gr00Config.TcGVL
{attribute 'Tc2GvlVarNames'}
VAR_GLOBAL CONSTANT
	tgGr00FieldbusMasterStartUp		:TIME := t#60s;					(* Maximal start time for the fieldbus master / Maximale startzeit für den Busmaster *)
	tgGr00PowerSupplyOn				:TIME := t#2s;						(* Delay to switch the power supply on *)
	tgGr00PowerSupplyOff				:TIME := t#1s;						(* Delay to switch the power supply off *)
	tgGr00AirPressureOnDelay			:TIME := t#1s;						(* Delay air pressure on *)
	tgGr00AirPressureDelay			:TIME := t#2s;						(* Delay air pressure present *)
	tgGr00AirPressureBuildUp			:TIME := t#20s;					(* Max time to building up the air pressure  / Maximale Zeit zum erreichen des Solldrucks *)
	tgGr00LightCurtainDelay			:TIME := t#1s;						(* After time light Curtain safe *)
	tgGr00TempErrorDelay			:TIME := t#5m;						(* Max delay time until the message turns to an error *)
	rgGr00AdsOverrideAcc				:REAL := 10.0;						(* Override accerlation per second / Override Beschleuingung pro sekunde *)
	rgGr00AdsOverrideDec			:REAL :=100.0;					(* Override decerlation per second / Override Verzögerung pro sekunde *)
	sgGr00MachineLifetimeFilePath		:STRING := 'C:\TwinCAT\Boot\';(* File path for machine life time *)
	sgGr00MachineLifetimeFileName	:STRING := 'mlt';					(* File name for machine life time *)
	sgGr00PrgPath					:STRING := 'C:\TwinCAT\Boot\';(* Program path e.g. '\Hard Disk\Riex\Recipe'*)
	sgGr00PrgName					:STRING := 'prg';					(* Recipe name e.g. 'default' *)
	sgGr00PrgSuffix					:STRING := 'riex';					(* Recipe suffix e.g. rcp *)
END_VAR

// ---- Global Variables/Config/GVL_Gr01Config.TcGVL
{attribute 'Tc2GvlVarNames'}
VAR_GLOBAL CONSTANT
	tgGr01ControllerOff					:TIME := t#10s;				(* Delay to switch the controller off *)
	tgGr01LightCurtainDelay				:TIME := t#1s;					(* After time light Curtain safe *)
	tgGr01MaxRefTime					:TIME := t#4m;					(* Maximum time after start reference until message in reference / Maximale Zeit von Starten der Referenbzfahr bis ende der Referenzfahrt *)

	rgGr01AdsOverrideAcc					:REAL := 10.0;					(* Override accerlation per second / Override Beschleuingung pro sekunde *)
	rgGr01AdsOverrideDec				:REAL :=100.0;				(* Override decerlation per second / Override Verzögerung pro sekunde *)

	sgGr01LifetimeFilePath					:STRING := 'C:\TwinCAT\Boot\';	(* File path for life time *)
	sgGr01LifetimeFileName				:STRING := 'lt1';				(* File name for life time *)

	rGr01PipeDiameterMin					:REAL := 160;					(* 6.625" Minimal pipe diameter *)
	rGr01PipeDiameterMax				:REAL := 770;					(* 30" Maximal pipe diameter *)

	(* Axis angle parameters *)
	udngGr01AxisAngleInc					:UDINT := 8192;	  			(* Increment value of axis angle pro path[INC] *)
	lrgGr01AxisAnglePath					:LREAL := 360.0;  				(* Path lenght of axis angle [deg] *)

	lrgGr01AngleAutoMax					:LREAL := 45;					(* Maximal angle to sawing in automatic mode *)

	(* Saw band parameters*)
	udngGr01SawbandInc					:UDINT := 18;	  				(* Increment value of saw band pro rotation [INC] *)
	lrgGr01SawbandDistance				:LREAL := 1602.21;  			(* Rotation distance of saw band  [mm] *)

	tgGr01SawbandAirOffDelay				:TIME := t#10s;				(* Sawband air off delay *)
	tgGr01VacuumCleanerOffDelay			:TIME := t#10s;				(* Vacuum cleaner off delay *)
	tgGr01SawbandReadyDelay			:TIME := t#5s;					(* Sawband ready delay *)
	tgGr01SpeedNoConstant		 		:TIME := t#3s;					(* Sawband speed no constant *)

END_VAR

// ---- Global Variables/Config/GVL_Gr02Config.TcGVL
{attribute 'Tc2GvlVarNames'}
VAR_GLOBAL CONSTANT
	tgGr02ControllerOff					:TIME := t#10s;				(* Delay to switch the controller off *)
	tgGr02LightCurtainDelay				:TIME := t#1s;					(* After time light Curtain safe *)
	tgGr02MaxRefTime					:TIME := t#4m;					(* Maximum time after start reference until message in reference / Maximale Zeit von Starten der Referenbzfahr bis ende der Referenzfahrt *)

	rgGr02AdsOverrideAcc					:REAL := 10.0;					(* Override accerlation per second / Override Beschleuingung pro sekunde *)
	rgGr02AdsOverrideDec				:REAL :=100.0;				(* Override decerlation per second / Override Verzögerung pro sekunde *)

	sgGr02LifetimeFilePath					:STRING := 'C:\TwinCAT\Boot\';	(* File path for saw band enabled life time *)
	sgGr02LifetimeFileName				:STRING := 'lt2';				(* File name for saw band enabled life time *)

	(* Axis parameters *)

END_VAR

// ---- Global Variables/Config/GVL_Gr05Config.TcGVL
{attribute 'Tc2GvlVarNames'}
VAR_GLOBAL CONSTANT
	tgGr05ControllerOff					:TIME := T#10S;				(* Delay to switch the controller off *)
	tgGr05LightCurtainDelay				:TIME := T#1S;					(* After time light Curtain safe *)
	tgGr05MaxRefTime					:TIME := T#4M;					(* Maximum time after start reference until message in reference / Maximale Zeit von Starten der Referenbzfahr bis ende der Referenzfahrt *)

	rgGr05AdsOverrideAcc				:REAL := 10.0;					(* Override accerlation per second / Override Beschleuingung pro sekunde *)
	rgGr05AdsOverrideDec				:REAL :=100.0;				(* Override decerlation per second / Override Verzögerung pro sekunde *)

	sgGr05LifetimeFilePath				:STRING := 'C:\TwinCAT\Boot\';	(* File path for life time *)
	sgGr05LifetimeFileName				:STRING := 'lt5';				(* File name for life time *)

	(* Clamp cylinder parameters *)
	ungGr05ClampMaxNo					:UINT := 2;					(* Maxinmal number of clamps *)

	(* Position cylinder parameters *)
	lrgGr05CylinderPosOffset			:LREAL := 100;				(* Position offset *)
	lrgGr05CylinderPosOriginShiftPos	:LREAL := 0;				(* Orgin shift position *)
	etgGr05CylinderPosDirection			:ET_MC_Direction := ET_MC_Direction_ePositive;				(* Direction: -1 Negative, +1 Positive *)
	usngGr05CylinderPosCodingType		:USINT := 1;
	ungGr05CylinderPosMaxNo				:UINT := 3;					(* Maxinmal number of position cylinders *)

	(* Spindle starting parameters *)
	ungGr05MaxPhasesNewSpdl 			:UINT := 4;					(* Max number of starting phases for new spindle *)
	ungGr05MaxPhasesDailyPreheat		:UINT := 4;					(* Max number of starting  phases for daily preheat *)
END_VAR

// ---- Global Variables/FB_Alarm/GVL_FB_Alarm.TcGVL
{attribute 'Tc2GvlVarNames'}
VAR_GLOBAL CONSTANT
	nALARM_MAX_NO			:INT := 31;			(* Maximal number of alarms *)
END_VAR

// ---- Global Variables/FB_Fieldbus/GVL_FB_Fieldbus.TcGVL
{attribute 'Tc2GvlVarNames'}
VAR_GLOBAL CONSTANT
	iSLAVEADDR_ARR_SIZE	: DINT := 256;
	dnDIAG_SLAVEINFO_SIZE	:DINT := 10;
END_VAR
VAR_GLOBAL
	SaveDiagSlaveInfo 			:ARRAY [0..dnDIAG_SLAVEINFO_SIZE] OF ST_SlaveStateInfo;
	SaveDiagSlaveInfoScanned	:ARRAY [0..dnDIAG_SLAVEINFO_SIZE] OF ST_SlaveStateInfoScanned;
END_VAR

// ---- Global Variables/FB_GFX4IRZones/GVL_FB_GFX4IRZones.TcGVL
{attribute 'Tc2GvlVarNames'}
VAR_GLOBAL CONSTANT
	nZONES_MAX_NO			:UINT := 4;			(* Amount of control zones *)
END_VAR

// ---- Global Variables/FB_LoadFromFile/GVL_FB_LoadFromFile.TcGVL
{attribute 'Tc2GvlVarNames'}
VAR_GLOBAL CONSTANT
	usnFileArrayMaxDimR					:USINT := 100;		(* 0..usnMaxDimR - Number of rows to read. *)
	usnFileArrayMaxDimC					:USINT := 1;  			(* 0..usnMaxDimC -  Number of columns to read. *)
END_VAR

// ---- Global Variables/FB_Logger/GVL_FB_Logger.TcGVL
{attribute 'Tc2GvlVarNames'}
VAR_GLOBAL
	unLOG_INSTANCE_IDX				:UINT;
END_VAR
VAR_GLOBAL CONSTANT
	sLOG_FILE_PATH					:STRING := '\Hard Disk\Riex\Log\';			(* Login file path *)
	sLOG_FILE_SUFFIX					:STRING := 'log';							(* Suffix of loggin file *)
	unNUM_OF_LOG_VAR					:UINT := 4;								(* Number of logging variables *)
	unLOG_MAX_NO						:UINT := 1;
	unLOG_BEFOR_MAX_NO				:UINT := 10;
	unLOG_DURING_MAX_NO				:UINT := 250;
	unLOG_AFTER_MAX_NO				:UINT := 10;
END_VAR

// ---- Global Variables/FB_Traceability/GVL_Traceability.TcGVL
{attribute 'Tc2GvlVarNames'}
VAR_GLOBAL CONSTANT
	bTraceEnable						:BOOL := TRUE;					(* Traceability enable *)
	sTracePath							:STRING := '\Hard Disk\Riex\Traceability\NewData\';	(* Path to file e.g. 'c:\', \Hard Disk\ *)
	sTraceFileName						:STRING(20);						(* Name of file *)
	sTraceFileExtension					:STRING(5) := 'txt';					(* File extension  *)
	sTraceColSep						:STRING(5) := '$T';					(* Seperator sign for columns *)
	udnTraceStringLengthMax 				:UDINT := 255;
	udnTraceSampleMax 					:UDINT := 101;
	udnTraceDataMax 					:UDINT := 19;
END_VAR

// ---- Global Variables/GVL.TcGVL
{attribute 'Tc2GvlVarNames'}
VAR_GLOBAL
	sgAmsNetId					:STRING := '';						(* AmsNetID of the controller, '' = local netid *)
	lrgActCycleTime				:LREAL;								(* Actual cycle time *)
	// stgSystemTaskInfoArr       		AT%MB32832 :ARRAY[1..4] OF SYSTEMTASKINFOTYPE;
	
	_PlcAppSystemInfo			:PlcAppSystemInfo;
	_PlcTaskSystemInfo			:PlcTaskSystemInfo;	
END_VAR

// ---- Global Variables/GVL_Gr0000.TcGVL
{attribute 'Tc2GvlVarNames'}
VAR_GLOBAL
	etgGr00MachineMode				:ET_MachineMode;			(* Machine mode *)
	etgGr00MachineState				:ET_MachineState;			(* Machine state *)
	stgGr00Blinker					:ST_Blinker;
	bgGr00NoEmergencyStop			:BOOL;						(* No ermergency Stop / Keine Notaus *)
	bgGr00AirPressureOK				:BOOL;						(* Air Pressure is available / Luftdruck ist vorhanden *)
	bgGr00LightCurtainOK				:BOOL;						(* Light curtain ok / Freigabe Lichtschranke i.o *)
	bgGr00PowerSupplyOk			:BOOL;						(* Power supply on / Leitung eingeschaltet *)
	bgGr00AllDoorsClosed				:BOOL;						(* All doors closed / Alle Türen geschlossen *)
	bgGr00AllDoorsClosedLocked		:BOOL;						(* All doors closed and locked / Alle Türen geschlossen und verrrigelt *)
	bgGr00ModeAutomatic				:BOOL;						(* Machine mode automatic *)
	bgGr00ModeHome				:BOOL;						(* Machine mode home *)
	bgGr00ModeManual				:BOOL;						(* Machine mode manual *)
	bgGr00MachineRunning			:BOOL;						(* Machine running / Maschine lauft *)
	bgGr00MachineStandstill			:BOOL;						(* Machine standstill / Maschin steht *)
	bgGr00SafetyCompleted			:BOOL;						(* Safety completed *)
	bgGr00ManualCompleted			:BOOL;						(* Manual completed *)
	bgGr00HomeCompleted			:BOOL;						(* Home completed / Grundsrellung ausgeführt *)
	bgGr00AutoCompleted				:BOOL;						(* Automatic completed / Automatik beendet *)
	bgGr00MoveInterrupted			:BOOL;						(* Move interrupted / Bewegung unterbrochen *)
	bgGr00ConfirmAlarm				:BOOL;						(* Confirm alarm *)
	bgGr00MachinePurge				:BOOL;						(* Machine purge *)
	rgGr00Override					:REAL;						(* Override *)
	bgGr00WritePersistent				:BOOL;						(* Write persisten data *)
	stgGr00DateTime					:ST_DateTime;				(* Current date and time *)
	bgGr00HomeNotInCrashGr01		:BOOL;						(* Home not in crash for Gr01 output *)
	arrGr00ProcessPara				:ARRAY [0..usnFileArrayMaxDimR, 0..usnFileArrayMaxDimC ] OF REAL; 			(* Matrix with process parameters from file *)
	bgGr00DoorsUnlockRequest 		:BOOL;						(* Doors unlock request *)
	bgGr00DoorsUnlockRelease		:BOOL;						(* Doors unlock release *)
END_VAR

// ---- Global Variables/GVL_Gr0100.TcGVL
{attribute 'Tc2GvlVarNames'}
VAR_GLOBAL
	arbgGr01StartProcess			:ARRAY[1..3] OF BOOL;		(* Start process *)
	bgGr01LightCurtainOK			:BOOL;						(* Light curtain ok / Freigabe Lichtschranke i.o *)
	bgGr01HomeNotInCrashGr02		:BOOL;						(* Home not in crash for Gr02 output *)
	bgGr01HomeNotInCrashGr05		:BOOL;						(* Home not in crash for Gr05 output *)
	bgGr01NotInCrashArea			:BOOL;						(* Axis not in crash are with *)
	bgGr01SafetyCompleted			:BOOL;						(* Safety completed *)
	bgGr01ManualCompleted			:BOOL;						(* Manual completed *)
	bgGr01HomeCompleted				:BOOL;						(* Home completed / Grundsrellung ausgeführt *)
	bgGr01AutoCompleted				:BOOL;						(* Automatic completed / Automatik beendet *)
	bgGr01MoveInterrupted			:BOOL;						(* Move interrupted / Bewegung unterbrochen *)
	bgGr01WritePersistent			:BOOL;						(* Write persisten data *)
	bgGr01SafetyActive				:BOOL;						(* Safety active *)
	bgGr01SawingAck 				:BOOL;						(* Ack from Gr01 to Gr05 *)
	bgGr01AngleAck					:BOOL;						(* Ack from Gr01 to Gr05 *)
	bgGr01TransportReq				:BOOL;						(* Req from Gr01 to Gr05 *)
	bgGr01PipePresent				:BOOL;						(* Pipe present *)
	
	bgGr01SawbandVeloError_1		:BOOL;						(* Sawband stand still *)
	bgGr01SawbandVeloError_2		:BOOL;						(* Sawband Velocity is to low *)
	bgGr01SawbandInSpeed			:BOOL;						(* Sawband is in speed *)
END_VAR

// ---- Global Variables/GVL_Gr0200.TcGVL
{attribute 'Tc2GvlVarNames'}
VAR_GLOBAL
	arbgGr02StartProcess				:ARRAY[1..3] OF BOOL;		(* Start process *)
	bgGr02LightCurtainOK				:BOOL;						(* Light curtain ok / Freigabe Lichtschranke i.o *)
	bgGr02HomeNotInCrashGr02		:BOOL;						(* Home not in crash for Gr02 output *)
	bgGr02HomeNotInCrashGr05		:BOOL;						(* Home not in crash for Gr05 output *)
	bgGr02NotInCrashArea				:BOOL;						(* Axis not in crash are with *)
	bgGr02SafetyCompleted			:BOOL := TRUE;				(* Safety completed *)
	bgGr02ManualCompleted			:BOOL := TRUE;				(* Manual completed *)
	bgGr02HomeCompleted			:BOOL := TRUE;				(* Home completed / Grundsrellung ausgeführt *)
	bgGr02AutoCompleted				:BOOL := TRUE;				(* Automatic completed / Automatik beendet *)
	bgGr02MoveInterrupted			:BOOL;						(* Move interrupted / Bewegung unterbrochen *)
	bgGr02WritePersistent				:BOOL;						(* Write persisten data *)
	bgGr02SafetyActive				:BOOL;						(* Safety active *)
END_VAR

// ---- Global Variables/GVL_Gr0500.TcGVL
{attribute 'Tc2GvlVarNames'}
VAR_GLOBAL
	bgGr05StartProcess				:BOOL;						(* Start process *)
	bgGr05LightCurtainOK				:BOOL;						(* Light curtain ok / Freigabe Lichtschranke i.o *)
	bgGr05HomeNotInCrashGr01		:BOOL;						(* Home not in crash for Gr01 output *)
	bgGr05HomeNotInCrashGr02		:BOOL;						(* Home not in crash for Gr02 output *)
	bgGr05SafetyCompleted			:BOOL;						(* Safety completed *)
	bgGr05ManualCompleted			:BOOL;						(* Manual completed *)
	bgGr05HomeCompleted			:BOOL;						(* Home completed / Grundsrellung ausgeführt *)
	bgGr05AutoCompleted				:BOOL;						(* Automatic completed / Automatik beendet *)
	bgGr05MoveInterrupted			:BOOL;						(* Move interrupted / Bewegung unterbrochen *)
	bgGr05WritePersistent				:BOOL;						(* Write persisten data *)
	bgGr05SafetyActive				:BOOL;						(* Safety active *)
	bgGr05SawingReq 				:BOOL;						(* Req from Gr05 to Gr01 *)
	bgGr05AngleReq 					:BOOL;						(* Req from Gr05 to Gr01 *)
	bgGr05TransportAck 				:BOOL;						(* Ack from Gr05 to Gr01 *)
	bgGr05PipeEndPresent			:BOOL;						(* End of pipe present *)
	bgGr05PipeBeginPresent			:BOOL;						(* Begin of pipe present *)
	lrgGr05SafetyDistance				:LREAL;						(* *)
END_VAR

// ---- Global Variables/HMI/GVL_Gr00HMI.TcGVL
{attribute 'Tc2GvlVarNames'}
VAR_GLOBAL
	stgGr00HMI			:ST_Gr00HMIRef;
END_VAR

// ---- Global Variables/HMI/GVL_Gr01HMI.TcGVL
{attribute 'Tc2GvlVarNames'}
VAR_GLOBAL
	stgGr01HMI			:ST_Gr01HMIRef;
END_VAR

// ---- Global Variables/HMI/GVL_Gr02HMI.TcGVL
{attribute 'Tc2GvlVarNames'}
VAR_GLOBAL
	stgGr02HMI			:ST_Gr02HMIRef;
END_VAR

// ---- Global Variables/HMI/GVL_Gr05HMI.TcGVL
{attribute 'Tc2GvlVarNames'}
VAR_GLOBAL
	stgGr05HMI			:ST_Gr05HMIRef;
END_VAR

// ---- Global Variables/Init/GVL_Gr00Init.TcGVL
{attribute 'Tc2GvlVarNames'}
VAR_GLOBAL
		tPLC_TaskCycleTime_ms			:TIME 	:=	LREAL_TO_TIME(GVL.lrgActCycleTime * 1000) ;		(* PLC Task Cycle Time in [ms] *)
END_VAR

// ---- Global Variables/Init/GVL_Gr01Init.TcGVL
{attribute 'Tc2GvlVarNames'}
VAR_GLOBAL
	lrgGr01SawingSpeed					:LREAL := 30.78;				(* Sawing speed where 100% = 20 [mm/s] *)
	lrgGr01SawingEndPosition			:LREAL := -1.0;					(* Sawing end postion [mm] *)
	lrgGr01SawingEndDelay				:TIME := t#0.5s;				(* Wait after sawing done *)

	lrgGr01DistSawbandPipe				:LREAL := 80.00;				(* Distance between sawband an pipe present sensor *)
	
	rRaddurchmesser_mm					:REAL := 510.0;					(* Raddurchmesser für Sägebandgeschwindigkeit *) 
	uiImpulsDiscAmount					:UINT := 18;					(* 18 impulses on disc *)
END_VAR

// ---- Global Variables/Init/GVL_Gr02Init.TcGVL
{attribute 'Tc2GvlVarNames'}
VAR_GLOBAL

END_VAR

// ---- Global Variables/Init/GVL_Gr05Init.TcGVL
{attribute 'Tc2GvlVarNames'}
VAR_GLOBAL
	lrgGr05Clamp1DistPipeBeginSawBand		:LREAL := 710.0;			(* Distance between Sensor [pipe begin] and saw band (CAD) *)
	lrgGr05SearchDistPipeBegin				:LREAL := 500.0;			(* Search distance for the pipe begin  *)
	lrgGr05SearchDistPipeEnd					:LREAL := 180;			(* Search distance for the pipe end for last cut. Leftover piece as a good part, rest is cut *)

	lrgGr05Clamp1PipeSensorOffset				:LREAL := 205.0;			(* Pipe sensor position on axis clamp 1 (CAD) *)

	lrgGr05Clamp2PipeBeginPos				:LREAL := 0.0;				(* Position for pipe begin sensor *)
	lrgGr05Clamp2SawPos						:LREAL := 0.0;				(* Sawing position *)
	lrgGr05Clamp2Width						:LREAL := 150.0;			(* Width of clamping 2 support  *)

	lrgGr05RemovalBandSawBand				:LREAL := 500.0;			(* Distance from removal band to saw band *)

	tgGr05SlideWaitInWork					:TIME := t#2s;				(* Slide wait in work *)

	lrgGr05PipeClampWidth 					:LREAL := 120.0;			(* Pipe clamp width *)
	lrgGr05SawbandGuideWidth				:LREAL := 100.0;			(* Sawband guide width *)

END_VAR

// ---- Global Variables/Interface/GVL_Gr00Interface.TcGVL
{attribute 'Tc2GvlVarNames'}
VAR_GLOBAL
	(* Periphery *)
	Periphery					:ST_PERIPHERY_REF;
	iAxisDummy					:AXIS_REF;
END_VAR

// ---- Global Variables/Interface/GVL_Gr01Interface.TcGVL
{attribute 'Tc2GvlVarNames'}
VAR_GLOBAL
	(* Old from Tc2)
	(* Axis interface *)
	igGr01AxisSawBow			:ST_AXIS_REF;							(* Interface of axis saw bow *)
	igGr01AxisAngle				:ST_AXIS_REF;							(* Interface of axis angle *)

	igGr01AxisSawband			:ST_AXIS_REF;							(* Interface of axis sawband *)

	(* Drive interface *)
	igGr01DriveSawBow			:ST_DRIVE_REF;							(* Interface of drive saw bow *)
	igGr01DriveAngle			:ST_DRIVE_REF;							(* Interface of drive angle *)

	igGr01DriveSawband			:ST_DRIVE_REF;							(* Interface of drive sawband *)
*)

	(* Axis Interface) 			*)
	igGr01AxisSawBow			:AXIS_REF;								(* Interface plc -> nc *)
	igGr01AxisSawAngle			:AXIS_REF;								(* Interface plc -> nc *)
	igGr01AxisSawBand			:AXIS_REF;								(* Interface plc -> nc *)	
	
	
	(* Drive Interface)			*)
	igGr01DriveSawBow			:ST_STOEBERSI6SC6CIA402_REF;			(* Interface nc -> plc *)
	igGr01DriveSawAngle			:ST_STOEBERSI6SC6CIA402_REF;			(* Interface nc -> plc *)
	igGr01DriveSawBand			:ST_STOEBERSI6SC6CIA402_REF;			(* Interface nc -> plc *)
	
END_VAR

// ---- Global Variables/Interface/GVL_Gr02Interface.TcGVL
{attribute 'Tc2GvlVarNames'}
VAR_GLOBAL

END_VAR

// ---- Global Variables/Interface/GVL_Gr05Interface.TcGVL
{attribute 'Tc2GvlVarNames'}
VAR_GLOBAL
	(* Axis interface *)
	igGr05AxisClamp1			:AXIS_REF;							(* Interface plc -> nc *)

	(* Drive interface *)
	igGr05DriveClamp1			:ST_STOEBERSI6SC6CIA402_REF;		(* Interface nc -> plc *)

END_VAR

// ---- Global Variables/IO/GVL_Gr00IO.TcGVL
{attribute 'Tc2GvlVarNames'}
VAR_GLOBAL
(* Inputs / Eingänge *)
	stinGr00FieldbusStatus					AT %I*:ST_FieldbusStatus;										(* 		State of the fieldbus / Status des Fieldbus *)

	binGr00NoEmergencyStop					AT %I*:BOOL;													(*) 	No emergency stop / kein Notaus *)
	binGr00AirPressureOK					AT %I*:BOOL;													(*) 	Air pressure OK / Luftdruck i.O. *)
	arbinGr00DoorsClosed					AT %I* :ARRAY [1..5] OF BOOL;									(*) 	Doors closed / Türe geschlossen *)
	arbinGr00PowerSupplyOn					AT %I* :ARRAY [1..5] OF BOOL;									(*) 	Power supply on / 24V DC vorhanden. *)
	binGr00LightCurtainOK					AT %I*:BOOL;													(*) 	Light curtain ok / Freigabe Lichtschranke i.o *)
	binGr00TempOK							AT %I*:BOOL;													(*) 	Temperature fuse OK / Temperatursicherung i.O. *)
	binGr00AllDoorsClosed					AT %I*:BOOL;													(*) 	All doors closed / Alle Türen geschlossen *)
	binGr00AllDoorsLocked					AT %I*:BOOL;													(*) 	All doors locked / Alle Türen verriegelt *)

	binGr00PushBtnStart						AT %I*:BOOL;													(* DI 0.5)	Push button "Start" / Taste "Start" *)
	binGr00PushBtnStop						AT %I*:BOOL;													(* DI 0.6)	Push button "Stop" / Taste "Stop" *)
	binGr00PushBtnHome						AT %I*:BOOL;													(* DI 0.7)	Push button "Home" / Taster"Grundstellung" *)
	binGr00PushBtnReset						AT %I*:BOOL;													(* DI )	Push button "Reset" / Taste "Reset" *)
	binGr00PushBtnRef						AT %I*:BOOL;													(*) 	Push button "Ref" / Taste "Ref" *)

	binGr00PS6A24Ready						AT %I*:BOOL;													(* DI 10.1 PS6A24 is Ready; Ready if true *)
	binGr00PS6A24Warning_1					AT %I*:BOOL;													(* DI 10.3 PS6A24 Warning 1; Warning active if false; close to overload *)	
	binGr00PS6A24Warning_2					AT %I*:BOOL;													(* DI 10.5 PS6A24 Warning 2; Warning active if false; one or more phases out *)
	
	binGr00Luetze_F1						AT %I*:BOOL;													(* DI 10.0 DC Fuse F1 error *)
	binGr00Luetze_F2						AT %I*:BOOL;													(* DI 10.0 DC Fuse F2 error *)
	binGr00Luetze_F3						AT %I*:BOOL;													(* DI 10.0 DC Fuse F3 error *)
	
	
	(* Outputs / Ausgänge *)
	boutGr00AirPressureOn					AT %Q*:BOOL;													(* DQ 101.0) 	Air pressure on / Luftdruck ein. *)
	boutGr00ConfLightCurtain				AT %Q*:BOOL;													(*) 	Confirm light Curtain / Quitt Lichtschrank *)

	boutGr00BulbBtnStart					AT %Q*:BOOL;													(* DQ 0.5) 	Signal button bulb "start" / Signallampe "Start" *)
	boutGr00BulbBtnStop						AT %Q*:BOOL;													(* DQ 0.6) 	Signal button bulb "stop" / Signallampe "Stop" *)
	boutGr00BulbBtnHome						AT %Q*:BOOL;													(* DQ 0.7) 	Signal button bulb "home" / Signallampe "Grundstellung" *)
	boutGr00BulbBtnReset					AT %Q*:BOOL;													(* DQ 0.3) 	Signal button bulb "reset" / Signallampe "Reset" *)
	boutGr00BulbBtnRef						AT %Q*:BOOL;													(*) 	Signal button bulb "ref" / Signallampe "Ref" *)

	boutGr00BulbGreen						AT %Q*:BOOL;													(*) 	Signal column bulb "automatic" / Signallampe "Automatik" *)
	boutGr00BulbRed							AT %Q*:BOOL;													(*) 	Signal column bulb "stop" or "error" / Signallampe "Stop" oder "Fehler" *)
	boutGr00BulbYellow						AT %Q*:BOOL;													(*) 	Signal column bulb "warning" OR "message" / Signallampe "Warnung" oder "Message" *)
	boutGr00BulbWhite						AT %Q*:BOOL;													(*) 	Signal column bulb "" / Signallampe "" *)
	boutGr00Horn							AT %Q*:BOOL;													(*) 	Signal horn / Signal hupe *)

	boutGr00AllDoorsLock					AT %Q*:BOOL;													(* DQ 10.2) 	All doors lock / Alle Türen verriegeln *)
	

END_VAR

// ---- Global Variables/IO/GVL_Gr01IO.TcGVL
{attribute 'Tc2GvlVarNames'}
VAR_GLOBAL
	(* Inputs / Eingänge *)
	binGr01LightCurtainOK 					AT %I*:BOOL;													(*)		Light curtain ok / Freigabe Lichtschranke i.o *)

	binGr01PushBtnStart 					AT %I*:BOOL; 													(*)		Push button "Start" / Taste "Start" *)
	binGr01PushBtnStop 						AT %I*:BOOL; 													(*)		Push button "Stop" / Taste "Stop" *)

	binGr01AxisSawBowLimitMax 				AT %I*:BOOL; 													(* DI 110.0) 	Maximum limit of saw bow axis / Endschalter Bügel- Achse maximal *)
	binGr01AxisSawBowLimitMin 				AT %I*:BOOL; 													(* DI 110.1) 	Minimum limit of saw bow axis / Endschalter Bügel- Achse minimal *)
	binGr01AxisAngleLimitMax 				AT %I*:BOOL; 													(* DI 109.1) 	Maximum limit of angle axis / Endschalter Winkel - Achse maximal *)
	binGr01AxisAngleLimitMin 				AT %I*:BOOL; 													(* DI 109.0) 	Minimum limit of angle axis / Endschalter Winkel - Achse minimal *)

	binGr01SawbandRelease					AT %I*:BOOL;													(* DI 102.0)		Saw band release / Sägeband-Freigabe *)
	binGr01SawbandLocked					AT %I*:BOOL;													(* DI 102.1)		Currently not active *)
	binGr01SawbandMotorNOK					AT %I*:BOOL;													(*) 	DIx.x Saw band motor protection switch is no ok / Sägeband-Motorschutzschalter NiO *)
	binGr01SawbandNoBroken					AT %I*:BOOL;													(*) 	DI2.6 Saw band brake / Sägebandbruch *)

	binGr01VacuumCleanerMotorNOK			AT %I*:BOOL; 													(*) 	DIx.x Vacuum cleaner motor protection switch is no ok / Absaugung-Motorschutzschalter NiO *)

	binGr01PipeNoIdentify					AT %I*:BOOL;													(* DI 106.0) 	DI100.1 Pipe identify  / Rohrerkenung *)

	udninGr01CounterSawbandSpeed			AT %I*:UDINT;													(*) 	Counter Saw band speed counter / Sägeband-Geschwindigkeits-Zähler *)
	udninGr01IncAxisAngle					AT %I*:UDINT;													(*) 	SSI01 Axis angle increment *)
	
	ninGr01SawingOverride					AT %I*:INT;														(*) 	Sawing override *)

	(* Outputs / Ausgänge *)
	boutGr01ConfLightCurtain 				AT %Q*:BOOL; 													(*) 	Confirm light Curtain / Quitt Lichtschrank *)

	boutGr01BulbBtnStart 					AT %Q*:BOOL; 													(*) 	Signal button bulb "start" / Signallampe "Start" *)
	boutGr01BulbBtnStop 					AT %Q*:BOOL; 													(*) 	Signal button bulb "stop" / Signallampe "Stop" *)

	boutGr01SawbandAirOn					AT %Q*:BOOL;													(* DQ 101.2) 	Saw band air on / Sägeband Druckluft ein *)
	boutGr01LaserOn							AT %Q*:BOOL;													(* DQ 100.2) 	Laser on / off / Laser ein / aus *)
	boutGr01VacuumCleanerOn					AT %Q*:BOOL;													(*) 	Vacuum cleaner on / off / Absaugung ein / aus *)

	boutGr01SawBowAngleZero	 				AT %Q*:BOOL;													(* DQ 100.1) 	Saw bow angle zerro, confirmed safety is needed *)

END_VAR

// ---- Global Variables/IO/GVL_Gr02IO.TcGVL
{attribute 'Tc2GvlVarNames'}
VAR_GLOBAL
(* Inputs / Eingänge *)
	binGr02LightCurtainOK					AT %I*:BOOL;													(*) 	Light curtain ok / Freigabe Lichtschranke i.o *)

	binGr02PushBtnStart						AT %I*:BOOL;													(*) 	Push button "Start" / Taste "Start" *)
	binGr02PushBtnStop						AT %I*:BOOL;													(*) 	Push button "Stop" / Taste "Stop" *)

	(* Outputs / Ausgänge *)
	boutGr02ConfLightCurtain				AT %Q*:BOOL;													(*) 	Confirm light Curtain / Quitt Lichtschrank *)

	boutGr02BulbBtnStart					AT %Q*:BOOL;													(*) 	Signal button bulb "start" / Signallampe "Start" *)
	boutGr02BulbBtnStop						AT %Q*:BOOL;													(*) 	Signal button bulb "stop" / Signallampe "Stop" *)

END_VAR

// ---- Global Variables/IO/GVL_Gr05IO.TcGVL
{attribute 'Tc2GvlVarNames'}
VAR_GLOBAL
(* Inputs / Eingänge *)
	binGr05LightCurtainOK					AT %I*:BOOL;													(*) 	Light curtain ok / Freigabe Lichtschranke i.o *)

	binGr05PushBtnStart						AT %I*:BOOL;													(*) 	Push button "Start" / Taste "Start" *)
	binGr05PushBtnStop						AT %I*:BOOL;													(*) 	Push button "Stop" / Taste "Stop" *)

	binGr05AxisClamp1LimitMax				AT %I*:BOOL;													(* DI 108.0) 	Max Limit of clamp 1 feed; also ref point set with lrOriginShiftPos from HMI *)
	binGr05AxisClamp1LimitMin				AT %I*:BOOL;													(* DI 108.1) 	Min Limit of clamp 1 feed *)

	binGr05SlideTop							AT %I*:BOOL;													(*) 	Valve opened slide / Ventil Rutsche geöffnet *)
	binGr05SlideBottom						AT %I*:BOOL;													(*) 	Valve closed slide / Ventil Rutsche geschlossen *)

	binGr05RemovalBandNOK					AT %I*:BOOL;													(*) 	Removal band error / Abtransportband Fehler *)
	binGr05RemovalBandInPlus				AT %I*:BOOL;													(*) 	Removal band in plus limit / Abtransportband Plusendlage *)
	binGr05PushBtnRemovalBandStart			AT %I*:BOOL;													(*) 	Push button removal band "Start" / Taste Abtransportband "Start" *)
	binGr05RemovalBandInMinus				AT %I*:BOOL;													(*) 	Removal band in minus limit / Abtransportband Minusendlage *)

	arbinGr05ClampOpened					AT %I*: ARRAY[1..ungGr05ClampMaxNo] OF BOOL;					(*) 	Valve opened clamp 1, 2 / Ventil Klemmung 1, 2 geöffnet *)
	arbinGr05ClampClosed					AT %I*: ARRAY[1..ungGr05ClampMaxNo] OF BOOL;					(*) 	Valve closed clamp 1, 2  / Ventil Klemmung 1, 2  geschlossen *)

	arbinGr05CylinderPosOpened				AT %I*: ARRAY[1..ungGr05CylinderPosMaxNo] OF BOOL;				(* DI 103.0; 104.0; 105.0) 	Valve Pos Home | 100mm^=[1] | 200mm^=[2] | 300mm^=[3] *)
	arbinGr05CylinderPosClosed				AT %I*: ARRAY[1..ungGr05CylinderPosMaxNo] OF BOOL;				(* DI 103.1; 104.1; 105.1) 	Valves Pos Work | 100mm^=[1] | 200mm^=[2] | 300mm^=[3] *)

	binGr05PipeEndEdge						AT %I*:BOOL;													(* DI 106.1) 	Pipe end edge  / Rohrendekante *)
	binGr05PipeBeginEdge					AT %I*:BOOL;													(* DI 107.1) 	Pipe begin edge  / Rohranfangkante *)

	(* Outputs / Ausgänge *)
	boutGr05ConfLightCurtain				AT %Q*:BOOL;													(*) 	Confirm light Curtain / Quitt Lichtschrank *)

	boutGr05BulbBtnStart					AT %Q*:BOOL;													(*) 	Signal button bulb "start" / Signallampe "Start" *)
	boutGr05BulbBtnStop						AT %Q*:BOOL;													(*) 	Signal button bulb "stop" / Signallampe "Stop" *)

	boutGr05SlideUp							AT %Q*:BOOL;													(*) 	Valve open slide / Ventil Rutsche öffnen *)
	boutGr05SlideDown						AT %Q*:BOOL;													(*) 	Valve close slide / Ventil Rutsche schlissen *)

	boutGr05RemovalBandToPlus				AT %Q*:BOOL;													(*) 	Move removal band in plus direction / Abtransportband in Plusrichtung *)
	boutGr05RemovalBandToMinus				AT %Q*:BOOL;													(*) 	Move removal band in minus direction / Abtransportband in Minusrichtung *)


	arboutGr05ClampOpen						AT %Q*: ARRAY[1..ungGr05ClampMaxNo] OF BOOL;					(* DQ 102.0; 102.2) Valve Clamping MOVE to HomePos | Clamp_1^=[1] | Clamp_2^=[2] *)
	arboutGr05ClampClose					AT %Q*: ARRAY[1..ungGr05ClampMaxNo] OF BOOL;					(* DQ 102.1; 102.2)	Valve Clamping MOVE to WorkPos | Clamp_1^=[1] | Clamp_2^=[2] *)

	arboutGr05CylinderPosOpen				AT %Q*: ARRAY[1..ungGr05CylinderPosMaxNo] OF BOOL;				(* DQ 103.0; 103.2; 104.0) 	Valve MOVE to Pos Home | 100mm^=[1] | 200mm^=[2] | 300mm^=[3] *)
	arboutGr05CylinderPosClose				AT %Q*: ARRAY[1..ungGr05CylinderPosMaxNo] OF BOOL;				(* DQ 103.1; 103.3; 104.1) 	Valve MOVE to Pos Work | 100mm^=[1] | 200mm^=[2] | 300mm^=[3] *)

END_VAR

// ---- Global Variables/TwinCAT_Import.TcGVL
{attribute 'Tc2GvlVarNames'}
(* Generated automatically by TwinCAT - do not edit manually! *)
VAR_GLOBAL
END_VAR

